{region 'Documentation'}
(*!
<summary>Selects literal stimuli, gates and findings for a named checkpoint.</summary>
*)
{endregion}
METHOD PRIVATE SelectStep : BOOL //! TRUE after selecting a supported script step and its literal expectations; FALSE reports an unknown step.
SelectStep := FALSE;
FIntegerFinding := E_Result.NotEvaluated;
FTextFinding := E_Result.NotEvaluated;
FWideTextFinding := E_Result.NotEvaluated;
FRealFinding := E_Result.NotEvaluated;
FLRealFinding := E_Result.NotEvaluated;
CASE FStep OF
    StepInitialReset:
        FTrace := TraceScalarHistory;
        FResetSubjects := TRUE;
        FSample := 10;
        FTextSample := '10';
        FWideTextSample := "10";
        FRealSample.Value := 10.0;
        FLRealSample.Value := 10.0;
        FIntegerEnable := TRUE;
        FIntegerResult := E_Result.NotEvaluated;
        FIntegerObservation := FALSE;
        FIntegerEvaluation := FALSE;
        FTextEnable := TRUE;
        FTextResult := E_Result.NotEvaluated;
        FTextObservation := FALSE;
        FTextEvaluation := FALSE;
        FWideTextEnable := TRUE;
        FWideTextResult := E_Result.NotEvaluated;
        FWideTextObservation := FALSE;
        FWideTextEvaluation := FALSE;
        FRealEnable := TRUE;
        FRealResult := E_Result.NotEvaluated;
        FRealObservation := FALSE;
        FRealEvaluation := FALSE;
        FLRealEnable := TRUE;
        FLRealResult := E_Result.NotEvaluated;
        FLRealObservation := FALSE;
        FLRealEvaluation := FALSE;
    StepInitialObservation:
        FTrace := TraceScalarHistory;
        FResetSubjects := FALSE;
        FSample := 10;
        FTextSample := '10';
        FWideTextSample := "10";
        FRealSample.Value := 10.0;
        FLRealSample.Value := 10.0;
        FIntegerEnable := TRUE;
        FIntegerResult := E_Result.NotEvaluated;
        FIntegerObservation := TRUE;
        FIntegerEvaluation := FALSE;
        FTextEnable := TRUE;
        FTextResult := E_Result.NotEvaluated;
        FTextObservation := TRUE;
        FTextEvaluation := FALSE;
        FWideTextEnable := TRUE;
        FWideTextResult := E_Result.NotEvaluated;
        FWideTextObservation := TRUE;
        FWideTextEvaluation := FALSE;
        FRealEnable := TRUE;
        FRealResult := E_Result.NotEvaluated;
        FRealObservation := TRUE;
        FRealEvaluation := FALSE;
        FLRealEnable := TRUE;
        FLRealResult := E_Result.NotEvaluated;
        FLRealObservation := TRUE;
        FLRealEvaluation := FALSE;
    StepEqualObservation:
        FTrace := TraceScalarHistory;
        FResetSubjects := FALSE;
        FSample := 10;
        FTextSample := '10';
        FWideTextSample := "10";
        FRealSample.Value := 10.0;
        FLRealSample.Value := 10.0;
        FIntegerEnable := TRUE;
        FIntegerResult := E_Result.Passed;
        FIntegerObservation := TRUE;
        FIntegerEvaluation := TRUE;
        FTextEnable := TRUE;
        FTextResult := E_Result.Passed;
        FTextObservation := TRUE;
        FTextEvaluation := TRUE;
        FWideTextEnable := TRUE;
        FWideTextResult := E_Result.Passed;
        FWideTextObservation := TRUE;
        FWideTextEvaluation := TRUE;
        FRealEnable := TRUE;
        FRealResult := E_Result.Passed;
        FRealObservation := TRUE;
        FRealEvaluation := TRUE;
        FLRealEnable := TRUE;
        FLRealResult := E_Result.Passed;
        FLRealObservation := TRUE;
        FLRealEvaluation := TRUE;
    StepChangedObservation:
        FTrace := TraceScalarHistory;
        FResetSubjects := FALSE;
        FSample := 11;
        FTextSample := '11';
        FWideTextSample := "11";
        FRealSample.Value := 11.0;
        FLRealSample.Value := 11.0;
        FIntegerEnable := TRUE;
        FIntegerResult := E_Result.Failed;
        FIntegerObservation := TRUE;
        FIntegerEvaluation := TRUE;
        FIntegerFinding := E_Result.Failed;
        FTextEnable := TRUE;
        FTextResult := E_Result.Failed;
        FTextObservation := TRUE;
        FTextEvaluation := TRUE;
        FTextFinding := E_Result.Failed;
        FWideTextEnable := TRUE;
        FWideTextResult := E_Result.Failed;
        FWideTextObservation := TRUE;
        FWideTextEvaluation := TRUE;
        FWideTextFinding := E_Result.Failed;
        FRealEnable := TRUE;
        FRealResult := E_Result.Failed;
        FRealObservation := TRUE;
        FRealEvaluation := TRUE;
        FRealFinding := E_Result.Failed;
        FLRealEnable := TRUE;
        FLRealResult := E_Result.Failed;
        FLRealObservation := TRUE;
        FLRealEvaluation := TRUE;
        FLRealFinding := E_Result.Failed;
    StepReturnToInitial:
        FTrace := TraceScalarHistory;
        FResetSubjects := FALSE;
        FSample := 10;
        FTextSample := '10';
        FWideTextSample := "10";
        FRealSample.Value := 10.0;
        FLRealSample.Value := 10.0;
        FIntegerEnable := TRUE;
        FIntegerResult := E_Result.Failed;
        FIntegerObservation := TRUE;
        FIntegerEvaluation := TRUE;
        FTextEnable := TRUE;
        FTextResult := E_Result.Failed;
        FTextObservation := TRUE;
        FTextEvaluation := TRUE;
        FWideTextEnable := TRUE;
        FWideTextResult := E_Result.Failed;
        FWideTextObservation := TRUE;
        FWideTextEvaluation := TRUE;
        FRealEnable := TRUE;
        FRealResult := E_Result.Failed;
        FRealObservation := TRUE;
        FRealEvaluation := TRUE;
        FLRealEnable := TRUE;
        FLRealResult := E_Result.Failed;
        FLRealObservation := TRUE;
        FLRealEvaluation := TRUE;
    StepReenableReset:
        FTrace := TraceReenableBaseline;
        FResetSubjects := TRUE;
        FSample := 10;
        FTextSample := '10';
        FWideTextSample := "10";
        FRealSample.Value := 10.0;
        FLRealSample.Value := 10.0;
        FIntegerEnable := TRUE;
        FIntegerResult := E_Result.NotEvaluated;
        FIntegerObservation := FALSE;
        FIntegerEvaluation := FALSE;
        FTextEnable := TRUE;
        FTextResult := E_Result.NotEvaluated;
        FTextObservation := FALSE;
        FTextEvaluation := FALSE;
        FWideTextEnable := TRUE;
        FWideTextResult := E_Result.NotEvaluated;
        FWideTextObservation := FALSE;
        FWideTextEvaluation := FALSE;
        FRealEnable := TRUE;
        FRealResult := E_Result.NotEvaluated;
        FRealObservation := FALSE;
        FRealEvaluation := FALSE;
        FLRealEnable := TRUE;
        FLRealResult := E_Result.NotEvaluated;
        FLRealObservation := FALSE;
        FLRealEvaluation := FALSE;
    StepReenableBaseline:
        FTrace := TraceReenableBaseline;
        FResetSubjects := FALSE;
        FSample := 10;
        FTextSample := '10';
        FWideTextSample := "10";
        FRealSample.Value := 10.0;
        FLRealSample.Value := 10.0;
        FIntegerEnable := TRUE;
        FIntegerResult := E_Result.NotEvaluated;
        FIntegerObservation := TRUE;
        FIntegerEvaluation := FALSE;
        FTextEnable := TRUE;
        FTextResult := E_Result.NotEvaluated;
        FTextObservation := TRUE;
        FTextEvaluation := FALSE;
        FWideTextEnable := TRUE;
        FWideTextResult := E_Result.NotEvaluated;
        FWideTextObservation := TRUE;
        FWideTextEvaluation := FALSE;
        FRealEnable := TRUE;
        FRealResult := E_Result.NotEvaluated;
        FRealObservation := TRUE;
        FRealEvaluation := FALSE;
        FLRealEnable := TRUE;
        FLRealResult := E_Result.NotEvaluated;
        FLRealObservation := TRUE;
        FLRealEvaluation := FALSE;
    StepBeforeDisable:
        FTrace := TraceReenableBaseline;
        FResetSubjects := FALSE;
        FSample := 10;
        FTextSample := '10';
        FWideTextSample := "10";
        FRealSample.Value := 10.0;
        FLRealSample.Value := 10.0;
        FIntegerEnable := TRUE;
        FIntegerResult := E_Result.Passed;
        FIntegerObservation := TRUE;
        FIntegerEvaluation := TRUE;
        FTextEnable := TRUE;
        FTextResult := E_Result.Passed;
        FTextObservation := TRUE;
        FTextEvaluation := TRUE;
        FWideTextEnable := TRUE;
        FWideTextResult := E_Result.Passed;
        FWideTextObservation := TRUE;
        FWideTextEvaluation := TRUE;
        FRealEnable := TRUE;
        FRealResult := E_Result.Passed;
        FRealObservation := TRUE;
        FRealEvaluation := TRUE;
        FLRealEnable := TRUE;
        FLRealResult := E_Result.Passed;
        FLRealObservation := TRUE;
        FLRealEvaluation := TRUE;
    StepDisabledChange:
        FTrace := TraceReenableBaseline;
        FResetSubjects := FALSE;
        FSample := 20;
        FTextSample := '20';
        FWideTextSample := "20";
        FRealSample.Value := 20.0;
        FLRealSample.Value := 20.0;
        FIntegerEnable := FALSE;
        FIntegerResult := E_Result.Passed;
        FIntegerObservation := FALSE;
        FIntegerEvaluation := FALSE;
        FTextEnable := FALSE;
        FTextResult := E_Result.Passed;
        FTextObservation := FALSE;
        FTextEvaluation := FALSE;
        FWideTextEnable := FALSE;
        FWideTextResult := E_Result.Passed;
        FWideTextObservation := FALSE;
        FWideTextEvaluation := FALSE;
        FRealEnable := FALSE;
        FRealResult := E_Result.Passed;
        FRealObservation := FALSE;
        FRealEvaluation := FALSE;
        FLRealEnable := FALSE;
        FLRealResult := E_Result.Passed;
        FLRealObservation := FALSE;
        FLRealEvaluation := FALSE;
    StepReenabledCapture:
        FTrace := TraceReenableBaseline;
        FResetSubjects := FALSE;
        FSample := 20;
        FTextSample := '20';
        FWideTextSample := "20";
        FRealSample.Value := 20.0;
        FLRealSample.Value := 20.0;
        FIntegerEnable := TRUE;
        FIntegerResult := E_Result.Passed;
        FIntegerObservation := TRUE;
        FIntegerEvaluation := FALSE;
        FTextEnable := TRUE;
        FTextResult := E_Result.Passed;
        FTextObservation := TRUE;
        FTextEvaluation := FALSE;
        FWideTextEnable := TRUE;
        FWideTextResult := E_Result.Passed;
        FWideTextObservation := TRUE;
        FWideTextEvaluation := FALSE;
        FRealEnable := TRUE;
        FRealResult := E_Result.Passed;
        FRealObservation := TRUE;
        FRealEvaluation := FALSE;
        FLRealEnable := TRUE;
        FLRealResult := E_Result.Passed;
        FLRealObservation := TRUE;
        FLRealEvaluation := FALSE;
    StepReenabledComparison:
        FTrace := TraceReenableBaseline;
        FResetSubjects := FALSE;
        FSample := 20;
        FTextSample := '20';
        FWideTextSample := "20";
        FRealSample.Value := 20.0;
        FLRealSample.Value := 20.0;
        FIntegerEnable := TRUE;
        FIntegerResult := E_Result.Passed;
        FIntegerObservation := TRUE;
        FIntegerEvaluation := TRUE;
        FTextEnable := TRUE;
        FTextResult := E_Result.Passed;
        FTextObservation := TRUE;
        FTextEvaluation := TRUE;
        FWideTextEnable := TRUE;
        FWideTextResult := E_Result.Passed;
        FWideTextObservation := TRUE;
        FWideTextEvaluation := TRUE;
        FRealEnable := TRUE;
        FRealResult := E_Result.Passed;
        FRealObservation := TRUE;
        FRealEvaluation := TRUE;
        FLRealEnable := TRUE;
        FLRealResult := E_Result.Passed;
        FLRealObservation := TRUE;
        FLRealEvaluation := TRUE;
    StepResetNewBaseline:
        FTrace := TraceResetBaseline;
        FResetSubjects := TRUE;
        FSample := 30;
        FTextSample := '30';
        FWideTextSample := "30";
        FRealSample.Value := 30.0;
        FLRealSample.Value := 30.0;
        FIntegerEnable := TRUE;
        FIntegerResult := E_Result.NotEvaluated;
        FIntegerObservation := FALSE;
        FIntegerEvaluation := FALSE;
        FTextEnable := TRUE;
        FTextResult := E_Result.NotEvaluated;
        FTextObservation := FALSE;
        FTextEvaluation := FALSE;
        FWideTextEnable := TRUE;
        FWideTextResult := E_Result.NotEvaluated;
        FWideTextObservation := FALSE;
        FWideTextEvaluation := FALSE;
        FRealEnable := TRUE;
        FRealResult := E_Result.NotEvaluated;
        FRealObservation := FALSE;
        FRealEvaluation := FALSE;
        FLRealEnable := TRUE;
        FLRealResult := E_Result.NotEvaluated;
        FLRealObservation := FALSE;
        FLRealEvaluation := FALSE;
    StepNewBaselineCapture:
        FTrace := TraceResetBaseline;
        FResetSubjects := FALSE;
        FSample := 30;
        FTextSample := '30';
        FWideTextSample := "30";
        FRealSample.Value := 30.0;
        FLRealSample.Value := 30.0;
        FIntegerEnable := TRUE;
        FIntegerResult := E_Result.NotEvaluated;
        FIntegerObservation := TRUE;
        FIntegerEvaluation := FALSE;
        FTextEnable := TRUE;
        FTextResult := E_Result.NotEvaluated;
        FTextObservation := TRUE;
        FTextEvaluation := FALSE;
        FWideTextEnable := TRUE;
        FWideTextResult := E_Result.NotEvaluated;
        FWideTextObservation := TRUE;
        FWideTextEvaluation := FALSE;
        FRealEnable := TRUE;
        FRealResult := E_Result.NotEvaluated;
        FRealObservation := TRUE;
        FRealEvaluation := FALSE;
        FLRealEnable := TRUE;
        FLRealResult := E_Result.NotEvaluated;
        FLRealObservation := TRUE;
        FLRealEvaluation := FALSE;
    StepNewBaselineComparison:
        FTrace := TraceResetBaseline;
        FResetSubjects := FALSE;
        FSample := 30;
        FTextSample := '30';
        FWideTextSample := "30";
        FRealSample.Value := 30.0;
        FLRealSample.Value := 30.0;
        FIntegerEnable := TRUE;
        FIntegerResult := E_Result.Passed;
        FIntegerObservation := TRUE;
        FIntegerEvaluation := TRUE;
        FTextEnable := TRUE;
        FTextResult := E_Result.Passed;
        FTextObservation := TRUE;
        FTextEvaluation := TRUE;
        FWideTextEnable := TRUE;
        FWideTextResult := E_Result.Passed;
        FWideTextObservation := TRUE;
        FWideTextEvaluation := TRUE;
        FRealEnable := TRUE;
        FRealResult := E_Result.Passed;
        FRealObservation := TRUE;
        FRealEvaluation := TRUE;
        FLRealEnable := TRUE;
        FLRealResult := E_Result.Passed;
        FLRealObservation := TRUE;
        FLRealEvaluation := TRUE;
    StepNaNReset:
        FTrace := TraceScalarNonFinite;
        FResetSubjects := TRUE;
        FSample := 10;
        FTextSample := '10';
        FWideTextSample := "10";
        FRealSample.Value := 10.0;
        FLRealSample.Value := 10.0;
        FIntegerEnable := FALSE;
        FIntegerResult := E_Result.NotEvaluated;
        FIntegerObservation := FALSE;
        FIntegerEvaluation := FALSE;
        FTextEnable := FALSE;
        FTextResult := E_Result.NotEvaluated;
        FTextObservation := FALSE;
        FTextEvaluation := FALSE;
        FWideTextEnable := FALSE;
        FWideTextResult := E_Result.NotEvaluated;
        FWideTextObservation := FALSE;
        FWideTextEvaluation := FALSE;
        FRealEnable := FALSE;
        FRealResult := E_Result.NotEvaluated;
        FRealObservation := FALSE;
        FRealEvaluation := FALSE;
        FLRealEnable := FALSE;
        FLRealResult := E_Result.NotEvaluated;
        FLRealObservation := FALSE;
        FLRealEvaluation := FALSE;
    StepNaNCapture:
        FTrace := TraceScalarNonFinite;
        FResetSubjects := FALSE;
        FRealSample.Bits := DWORD#16#7FC00000;
        FLRealSample.Bits := LWORD#16#7FF8000000000000;
        FIntegerEnable := FALSE;
        FIntegerResult := E_Result.NotEvaluated;
        FIntegerObservation := FALSE;
        FIntegerEvaluation := FALSE;
        FTextEnable := FALSE;
        FTextResult := E_Result.NotEvaluated;
        FTextObservation := FALSE;
        FTextEvaluation := FALSE;
        FWideTextEnable := FALSE;
        FWideTextResult := E_Result.NotEvaluated;
        FWideTextObservation := FALSE;
        FWideTextEvaluation := FALSE;
        FRealEnable := TRUE;
        FRealResult := E_Result.Error;
        FRealObservation := TRUE;
        FRealEvaluation := FALSE;
        FRealFinding := E_Result.Error;
        FLRealEnable := TRUE;
        FLRealResult := E_Result.Error;
        FLRealObservation := TRUE;
        FLRealEvaluation := FALSE;
        FLRealFinding := E_Result.Error;
    StepNaNRepeated:
        FTrace := TraceScalarNonFinite;
        FResetSubjects := FALSE;
        // The same non-finite input must not produce duplicate findings.
        FIntegerEnable := FALSE;
        FIntegerResult := E_Result.NotEvaluated;
        FIntegerObservation := FALSE;
        FIntegerEvaluation := FALSE;
        FTextEnable := FALSE;
        FTextResult := E_Result.NotEvaluated;
        FTextObservation := FALSE;
        FTextEvaluation := FALSE;
        FWideTextEnable := FALSE;
        FWideTextResult := E_Result.NotEvaluated;
        FWideTextObservation := FALSE;
        FWideTextEvaluation := FALSE;
        FRealEnable := TRUE;
        FRealResult := E_Result.Error;
        FRealObservation := TRUE;
        FRealEvaluation := TRUE;
        FLRealEnable := TRUE;
        FLRealResult := E_Result.Error;
        FLRealObservation := TRUE;
        FLRealEvaluation := TRUE;
    StepPositiveInfinityReset:
        FTrace := TraceScalarNonFinite;
        FResetSubjects := TRUE;
        FSample := 10;
        FTextSample := '10';
        FWideTextSample := "10";
        FRealSample.Value := 10.0;
        FLRealSample.Value := 10.0;
        FIntegerEnable := FALSE;
        FIntegerResult := E_Result.NotEvaluated;
        FIntegerObservation := FALSE;
        FIntegerEvaluation := FALSE;
        FTextEnable := FALSE;
        FTextResult := E_Result.NotEvaluated;
        FTextObservation := FALSE;
        FTextEvaluation := FALSE;
        FWideTextEnable := FALSE;
        FWideTextResult := E_Result.NotEvaluated;
        FWideTextObservation := FALSE;
        FWideTextEvaluation := FALSE;
        FRealEnable := FALSE;
        FRealResult := E_Result.NotEvaluated;
        FRealObservation := FALSE;
        FRealEvaluation := FALSE;
        FLRealEnable := FALSE;
        FLRealResult := E_Result.NotEvaluated;
        FLRealObservation := FALSE;
        FLRealEvaluation := FALSE;
    StepPositiveInfinityCapture:
        FTrace := TraceScalarNonFinite;
        FResetSubjects := FALSE;
        FRealSample.Bits := DWORD#16#7F800000;
        FLRealSample.Bits := LWORD#16#7FF0000000000000;
        FIntegerEnable := FALSE;
        FIntegerResult := E_Result.NotEvaluated;
        FIntegerObservation := FALSE;
        FIntegerEvaluation := FALSE;
        FTextEnable := FALSE;
        FTextResult := E_Result.NotEvaluated;
        FTextObservation := FALSE;
        FTextEvaluation := FALSE;
        FWideTextEnable := FALSE;
        FWideTextResult := E_Result.NotEvaluated;
        FWideTextObservation := FALSE;
        FWideTextEvaluation := FALSE;
        FRealEnable := TRUE;
        FRealResult := E_Result.Error;
        FRealObservation := TRUE;
        FRealEvaluation := FALSE;
        FRealFinding := E_Result.Error;
        FLRealEnable := TRUE;
        FLRealResult := E_Result.Error;
        FLRealObservation := TRUE;
        FLRealEvaluation := FALSE;
        FLRealFinding := E_Result.Error;
    StepPositiveInfinityRepeated:
        FTrace := TraceScalarNonFinite;
        FResetSubjects := FALSE;
        // The same non-finite input must not produce duplicate findings.
        FIntegerEnable := FALSE;
        FIntegerResult := E_Result.NotEvaluated;
        FIntegerObservation := FALSE;
        FIntegerEvaluation := FALSE;
        FTextEnable := FALSE;
        FTextResult := E_Result.NotEvaluated;
        FTextObservation := FALSE;
        FTextEvaluation := FALSE;
        FWideTextEnable := FALSE;
        FWideTextResult := E_Result.NotEvaluated;
        FWideTextObservation := FALSE;
        FWideTextEvaluation := FALSE;
        FRealEnable := TRUE;
        FRealResult := E_Result.Error;
        FRealObservation := TRUE;
        FRealEvaluation := TRUE;
        FLRealEnable := TRUE;
        FLRealResult := E_Result.Error;
        FLRealObservation := TRUE;
        FLRealEvaluation := TRUE;
    StepNegativeInfinityReset:
        FTrace := TraceScalarNonFinite;
        FResetSubjects := TRUE;
        FSample := 10;
        FTextSample := '10';
        FWideTextSample := "10";
        FRealSample.Value := 10.0;
        FLRealSample.Value := 10.0;
        FIntegerEnable := FALSE;
        FIntegerResult := E_Result.NotEvaluated;
        FIntegerObservation := FALSE;
        FIntegerEvaluation := FALSE;
        FTextEnable := FALSE;
        FTextResult := E_Result.NotEvaluated;
        FTextObservation := FALSE;
        FTextEvaluation := FALSE;
        FWideTextEnable := FALSE;
        FWideTextResult := E_Result.NotEvaluated;
        FWideTextObservation := FALSE;
        FWideTextEvaluation := FALSE;
        FRealEnable := FALSE;
        FRealResult := E_Result.NotEvaluated;
        FRealObservation := FALSE;
        FRealEvaluation := FALSE;
        FLRealEnable := FALSE;
        FLRealResult := E_Result.NotEvaluated;
        FLRealObservation := FALSE;
        FLRealEvaluation := FALSE;
    StepNegativeInfinityCapture:
        FTrace := TraceScalarNonFinite;
        FResetSubjects := FALSE;
        FRealSample.Bits := DWORD#16#FF800000;
        FLRealSample.Bits := LWORD#16#FFF0000000000000;
        FIntegerEnable := FALSE;
        FIntegerResult := E_Result.NotEvaluated;
        FIntegerObservation := FALSE;
        FIntegerEvaluation := FALSE;
        FTextEnable := FALSE;
        FTextResult := E_Result.NotEvaluated;
        FTextObservation := FALSE;
        FTextEvaluation := FALSE;
        FWideTextEnable := FALSE;
        FWideTextResult := E_Result.NotEvaluated;
        FWideTextObservation := FALSE;
        FWideTextEvaluation := FALSE;
        FRealEnable := TRUE;
        FRealResult := E_Result.Error;
        FRealObservation := TRUE;
        FRealEvaluation := FALSE;
        FRealFinding := E_Result.Error;
        FLRealEnable := TRUE;
        FLRealResult := E_Result.Error;
        FLRealObservation := TRUE;
        FLRealEvaluation := FALSE;
        FLRealFinding := E_Result.Error;
    StepNegativeInfinityRepeated:
        FTrace := TraceScalarNonFinite;
        FResetSubjects := FALSE;
        // The same non-finite input must not produce duplicate findings.
        FIntegerEnable := FALSE;
        FIntegerResult := E_Result.NotEvaluated;
        FIntegerObservation := FALSE;
        FIntegerEvaluation := FALSE;
        FTextEnable := FALSE;
        FTextResult := E_Result.NotEvaluated;
        FTextObservation := FALSE;
        FTextEvaluation := FALSE;
        FWideTextEnable := FALSE;
        FWideTextResult := E_Result.NotEvaluated;
        FWideTextObservation := FALSE;
        FWideTextEvaluation := FALSE;
        FRealEnable := TRUE;
        FRealResult := E_Result.Error;
        FRealObservation := TRUE;
        FRealEvaluation := TRUE;
        FLRealEnable := TRUE;
        FLRealResult := E_Result.Error;
        FLRealObservation := TRUE;
        FLRealEvaluation := TRUE;
ELSE
    Error(Message := 'Unknown observation checkpoint.');
    RETURN;
END_CASE;
SelectStep := TRUE;
END_METHOD

END_FUNCTION_BLOCK

// ---- Framework/Assertions/POU/BasicTypes/DInt/AssertNoValueChange_DInt.TcPOU
{region 'Documentation'}
(*!
<summary>Check equality between consecutive active observations.</summary>
<description>

The first active observation establishes a baseline without deciding a result. Disabling
observation invalidates that baseline, not the held Result. Re-enabling first establishes a new
baseline; Reset clears history.

ObserveFirstCycle FALSE delays the first observation by one enabled call.

</description>
*)
{endregion}
FUNCTION_BLOCK AssertNoValueChange_DInt EXTENDS AssertionBase
VAR_INPUT
    IN : DINT; //! Actual value to observe.
END_VAR
VAR
    FINPrevious : DINT;
    FObservationPrevious : BOOL;
    FEvaluationActive : BOOL;
END_VAR

SUPER^();

{region 'Documentation'}
(*!
<summary>Observe the current value before evaluating a change against the previous observation.</summary>
*)
{endregion}
METHOD PROTECTED Assert
VAR
    PreviousValue : DINT;
    Message : STRING(GVL_Constants.MessageLength);
    PreviousText : STRING(GVL_Constants.AssertionValueLength);
    ActualText : STRING(GVL_Constants.AssertionValueLength);
END_VAR
FEvaluationActive := ObservationActive AND FObservationPrevious;
FObservationPrevious := ObservationActive;

IF NOT ObservationActive THEN
    RETURN;
END_IF;

PreviousValue := FINPrevious;
FINPrevious := IN;

IF NOT EvaluationActive THEN
    RETURN;
END_IF;

IF Result = E_Result.Error THEN
    RETURN;
END_IF;

IF Result = E_Result.Failed THEN
    RETURN;
END_IF;

IF IN <> PreviousValue THEN
    PreviousText := DINT_TO_STRING(PreviousValue);
    ActualText := DINT_TO_STRING(IN);
    Message := CONCAT('Assertion failed: value changed unexpectedly. Previous = ',
        PreviousText);
    Message := CONCAT(Message, ', Actual = ');
    Message := CONCAT(Message, ActualText);
    Message := CONCAT(Message, '.');
    Fail(Message := Message);
    RETURN;
END_IF;

Pass();
END_METHOD

{region 'Documentation'}
(*!
<summary>Current/last call has an active observation and a preceding observation
baseline.</summary>
*)
{endregion}
{attribute 'monitoring' := 'call'}
PROPERTY PUBLIC EvaluationActive : BOOL //! Current/last call has an active observation and a preceding observation baseline.
GET // PUBLIC
EvaluationActive := FEvaluationActive;
END_GET
END_PROPERTY

{region 'Documentation'}
(*!
<summary>Clear observation history and the current evaluation gate.</summary>
*)
{endregion}
METHOD PROTECTED ResetAssertion
FINPrevious := 0;
FObservationPrevious := FALSE;
FEvaluationActive := FALSE;
END_METHOD

END_FUNCTION_BLOCK

// ---- Framework/Assertions/POU/BasicTypes/LReal/AssertNoValueChange_LReal.TcPOU
{region 'Documentation'}
(*!
<summary>Check equality between consecutive active observations.</summary>
<description>

The first active observation establishes a baseline without deciding a result. Disabling
observation invalidates that baseline, not the held Result. Re-enabling first establishes a new
baseline; Reset clears history.

ObserveFirstCycle FALSE delays the first observation by one enabled call.

NaN or either infinity reports Error on an active observation, including baseline
capture; finite values compare exactly.

Numeric diagnostics use the formatter's default six significant digits; rounding affects
the message only, not the comparison.

</description>
*)
{endregion}
FUNCTION_BLOCK AssertNoValueChange_LReal EXTENDS AssertionBase
VAR_INPUT
    IN : LREAL; //! Actual value to observe.
END_VAR
VAR
    FINPrevious : LREAL;
    FObservationPrevious : BOOL;
    FEvaluationActive : BOOL;
END_VAR

SUPER^();

{region 'Documentation'}
(*!
<summary>Observe the current value before evaluating a change against the previous observation.</summary>
*)
{endregion}
METHOD PROTECTED Assert
VAR
    PreviousValue : LREAL;
    Message : STRING(GVL_Constants.MessageLength);
    PreviousText : STRING(GVL_Constants.AssertionValueLength);
    ActualText : STRING(GVL_Constants.AssertionValueLength);
END_VAR
FEvaluationActive := ObservationActive AND FObservationPrevious;
FObservationPrevious := ObservationActive;

IF NOT ObservationActive THEN
    RETURN;
END_IF;

PreviousValue := FINPrevious;
FINPrevious := IN;

IF Result = E_Result.Error THEN
    RETURN;
END_IF;

IF NOT Tc2_Utilities.LrealIsFinite(x := IN) THEN
    Error(Message := 'Assertion error: IN must be finite.');
    RETURN;
END_IF;

IF NOT EvaluationActive THEN
    RETURN;
END_IF;

IF Result = E_Result.Failed THEN
    RETURN;
END_IF;

IF IN <> PreviousValue THEN
    PreviousText := CreateAssertionTextValue_LReal(Value := PreviousValue);
    ActualText := CreateAssertionTextValue_LReal(Value := IN);
    Message := CONCAT('Assertion failed: value changed unexpectedly. Previous = ',
        PreviousText);
    Message := CONCAT(Message, ', Actual = ');
    Message := CONCAT(Message, ActualText);
    Message := CONCAT(Message, '.');
    Fail(Message := Message);
    RETURN;
END_IF;

Pass();
END_METHOD

{region 'Documentation'}
(*!
<summary>Current/last call has an active observation and a preceding observation
baseline.</summary>
*)
{endregion}
{attribute 'monitoring' := 'call'}
PROPERTY PUBLIC EvaluationActive : BOOL //! Current/last call has an active observation and a preceding observation baseline.
GET // PUBLIC
EvaluationActive := FEvaluationActive;
END_GET
END_PROPERTY

{region 'Documentation'}
(*!
<summary>Clear observation history and the current evaluation gate.</summary>
*)
{endregion}
METHOD PROTECTED ResetAssertion
FINPrevious := 0.0;
FObservationPrevious := FALSE;
FEvaluationActive := FALSE;
END_METHOD

END_FUNCTION_BLOCK

// ---- SelfTests/TestCases/TestSuite_AssertionObservation/Test_AssertionArraySnapshot.TcPOU
{region 'Documentation'}
(*!
<summary>Checks retained DINT array snapshots, independent bounds and delayed observation.</summary>
<description>
IN[-2..1] selects [-1..0], while Memory[5..7] stores two values and an untouched
tail sentinel. Disable never replaces the snapshot. Reset invalidates it without
clearing Memory; ObserveFirstCycle=FALSE delays capture until the second enabled
call. Literal memory checks distinguish fixed snapshots from rolling history.
Each named step calls each subject once and checks public gates, result and local
findings before advancing in the next cycle. Outer Assertions collect checkpoints
per trace; subjects never contribute their intentional failures to the test result.
FirstFailedStep retains the first mismatch. No timed stimulus or expected-result
algorithm is used.
</description>
*)
{endregion}
FUNCTION_BLOCK Test_AssertionArraySnapshot EXTENDS TestCaseBase
VAR
    FImmediate : AssertArrayNoValueChange_DInt;
    FDelayed : AssertArrayNoValueChange_DInt;
    FInput : ARRAY[-2..1] OF DINT;
    FImmediateMemory : ARRAY[5..7] OF DINT;
    FDelayedMemory : ARRAY[5..7] OF DINT;
    FExpectedImmediateFirst : DINT;
    FExpectedImmediateSecond : DINT;
    FExpectedDelayedFirst : DINT;
    FExpectedDelayedSecond : DINT;
    FCapture : EventBuffer;
    FEvents : ARRAY[1..CaptureLength] OF ST_Event;
    FCaptureFifo : ST_FifoStatus;
    FCaptureStatus : ST_EventBufferStatus;
    FSetupValid : BOOL;
    FStep : UINT;
    FTrace : UINT;
    FFirstFailedStep : UINT;
    FChecked : BOOL;
    FObservationReady : BOOL;
    FStepMatches : BOOL;
    FResultsMatch : BOOL;
    FActivityMatches : BOOL;
    FFindingsMatch : BOOL;
    FMemoryMatches : BOOL;
    FResetSubjects : BOOL;
    FImmediateEnable : BOOL;
    FImmediateResult : E_Result;
    FImmediateObservation : BOOL;
    FImmediateEvaluation : BOOL;
    FImmediateFinding : E_Result;
    FDelayedEnable : BOOL;
    FDelayedResult : E_Result;
    FDelayedObservation : BOOL;
    FDelayedEvaluation : BOOL;
    FDelayedFinding : E_Result;
    FFixedSnapshot : AssertTrue;
    FRetainedOnReenable : AssertTrue;
    FRecaptureAfterReset : AssertTrue;
END_VAR
VAR CONSTANT
    CaptureLength : UINT := 8;
    StepResetSnapshot : UINT := 1;
    StepFirstObservation : UINT := 2;
    StepDelayedCapture : UINT := 3;
    StepEqualSnapshot : UINT := 4;
    StepDivergence : UINT := 5;
    StepReturnToSnapshot : UINT := 6;
    StepResetForReenable : UINT := 7;
    StepReenableTraceCapture : UINT := 8;
    StepReenableTraceDelayedCapture : UINT := 9;
    StepReenableTracePassed : UINT := 10;
    StepDisabledChange : UINT := 11;
    StepReenableHistory : UINT := 12;
    StepReenableComparison : UINT := 13;
    StepReenableDelayedComparison : UINT := 14;
    StepResetKeepsMemory : UINT := 15;
    StepNewSnapshot : UINT := 16;
    StepNewDelayedSnapshot : UINT := 17;
    StepNewSnapshotMatches : UINT := 18;
    LastStep : UINT := StepNewSnapshotMatches;
    TraceFixedSnapshot : UINT := 1;
    TraceRetainedOnReenable : UINT := 2;
    TraceRecaptureAfterReset : UINT := 3;
END_VAR

SUPER^();

{region 'Documentation'}
(*!
<summary>Aggregates only the outer checks, not the intentionally failing subjects.</summary>
*)
{endregion}
METHOD PROTECTED AggregateResults
VAR_INPUT
    Aggregator : I_ResultAggregator; //! Borrowed result sink owned by the outer Test Case; add this test's checking Assertions without resetting or retaining the sink.
END_VAR
Aggregator.AddProvider(Provider := FFixedSnapshot);
Aggregator.AddProvider(Provider := FRetainedOnReenable);
Aggregator.AddProvider(Provider := FRecaptureAfterReset);
END_METHOD

{region 'Documentation'}
(*!
<summary>Calls each production subject with stable bindings and the selected stimulus.</summary>
*)
{endregion}
METHOD PRIVATE CallSubjects
FImmediate(Enable := FImmediateEnable,
    State := E_State.Running,
    StartIndex := -1,
    Length := 2,
    IN := FInput,
    Memory := FImmediateMemory);
FDelayed(Enable := FDelayedEnable,
    State := E_State.Running,
    StartIndex := -1,
    Length := 2,
    IN := FInput,
    Memory := FDelayedMemory);
END_METHOD

{region 'Documentation'}
(*!
<summary>Checks finding order, identities and exact count without retaining prior events.</summary>
*)
{endregion}
METHOD PRIVATE CheckFindings
VAR
    Index : UINT;
    FindingMatches : BOOL;
END_VAR
Index := 1;
FFindingsMatch := TRUE;
IF FImmediateFinding <> E_Result.NotEvaluated THEN
    FindingMatches := IsFindingValid(Index := Index,
        ExpectedName := FImmediate.Name,
        ExpectedResult := FImmediateFinding);
    FFindingsMatch := FFindingsMatch AND FindingMatches;
    Index := Index + 1;
END_IF;
IF FDelayedFinding <> E_Result.NotEvaluated THEN
    FindingMatches := IsFindingValid(Index := Index,
        ExpectedName := FDelayed.Name,
        ExpectedResult := FDelayedFinding);
    FFindingsMatch := FFindingsMatch AND FindingMatches;
    Index := Index + 1;
END_IF;
FFindingsMatch := FFindingsMatch
    AND (FCaptureStatus.SequenceId = UINT_TO_UDINT(Index - 1))
    AND (FCaptureStatus.LostEventCount = 0);
END_METHOD

{region 'Documentation'}
(*!
<summary>Rejects an incomplete capture or subject setup.</summary>
*)
{endregion}
METHOD PROTECTED CheckInitialization : BOOL //! TRUE when the inherited initialization check and this concrete fixture check both accept the setup.
CheckInitialization := SUPER^.CheckInitialization();
IF NOT CheckInitialization THEN
    RETURN;
END_IF;

CheckInitialization := FSetupValid
    AND FFixedSnapshot.IsInitialized
    AND FRetainedOnReenable.IsInitialized
    AND FRecaptureAfterReset.IsInitialized;
IF NOT CheckInitialization THEN
    EventPublisher.PublishEvent(Event := CreateFrameworkEvent(Name := Name,
        ResourceName := '',
        State := State,
        Severity := E_EventSeverity.Error,
        Message := 'Observation selftest setup failed.'));
END_IF;
END_METHOD

{region 'Documentation'}
(*!
<summary>Checks the selected snapshot and untouched sentinels.</summary>
*)
{endregion}
METHOD PRIVATE CheckMemory
FMemoryMatches := (FImmediateMemory[5] = FExpectedImmediateFirst)
    AND (FImmediateMemory[6] = FExpectedImmediateSecond)
    AND (FDelayedMemory[5] = FExpectedDelayedFirst)
    AND (FDelayedMemory[6] = FExpectedDelayedSecond)
    AND (FImmediateMemory[7] = -999)
    AND (FDelayedMemory[7] = -999)
    AND (FInput[-2] = -100)
    AND (FInput[1] = 100);
END_METHOD

{region 'Documentation'}
(*!
<summary>Checks literal result and observation/evaluation expectations.</summary>
*)
{endregion}
METHOD PRIVATE CheckResults
FResultsMatch := (FImmediate.Result = FImmediateResult)
    AND (FDelayed.Result = FDelayedResult);
FActivityMatches := (FImmediate.Enabled = FImmediateEnable)
    AND (FImmediate.ObservationActive = FImmediateObservation)
    AND (FImmediate.EvaluationActive = FImmediateEvaluation)
    AND (FDelayed.Enabled = FDelayedEnable)
    AND (FDelayed.ObservationActive = FDelayedObservation)
    AND (FDelayed.EvaluationActive = FDelayedEvaluation);
END_METHOD

{region 'Documentation'}
(*!
<summary>Initializes outer checks and isolates intentional subject findings.</summary>
*)
{endregion}
METHOD PROTECTED Configure
VAR
    Initialized : BOOL;
END_VAR
FPreparationStateCount := 0;
FTestStateCount := 1;
FFixedSnapshot.Initialize(Parent := THIS^,
    AssertionName := 'FixedSnapshot');
FRetainedOnReenable.Initialize(Parent := THIS^,
    AssertionName := 'RetainedOnReenable');
FRecaptureAfterReset.Initialize(Parent := THIS^,
    AssertionName := 'RecaptureAfterReset');
FSetupValid := FCapture.Initialize(Buffer := FEvents,
    FifoControl := FCaptureFifo,
    Status := FCaptureStatus);
FImmediate.BindPublisher(Publisher := FCapture);
Initialized := FImmediate.Initialize(Parent := THIS^,
    AssertionName := 'Immediate',
    ObserveFirstCycle := TRUE);
FSetupValid := FSetupValid AND Initialized;
FDelayed.BindPublisher(Publisher := FCapture);
Initialized := FDelayed.Initialize(Parent := THIS^,
    AssertionName := 'Delayed',
    ObserveFirstCycle := FALSE);
FSetupValid := FSetupValid AND Initialized;
END_METHOD

{region 'Documentation'}
(*!
<summary>Checks one expected Failed or Error finding from the bounded local capture.</summary>
*)
{endregion}
METHOD PRIVATE IsFindingValid : BOOL //! TRUE when the selected captured finding satisfies the scenario metadata and diagnostic checks.
VAR_INPUT
    Index : UINT; //! One-based index in the retained isolated event capture.
    ExpectedName : STRING(GVL_Constants.NameLength); //! Independently authored Assertion name expected in the selected finding.
    ExpectedResult : E_Result; //! Independently authored finding result.
END_VAR
IsFindingValid := (FEvents[Index].SequenceId = UINT_TO_UDINT(Index))
    AND (FEvents[Index].Name = ExpectedName)
    AND (FEvents[Index].OwnerScope = E_OwnerScope.Assertion)
    AND (FEvents[Index].EventType = E_EventType.Result)
    AND (FEvents[Index].State = E_State.Running)
    AND (FEvents[Index].Result = ExpectedResult)
    AND (FEvents[Index].Message <> '');
END_METHOD

{region 'Documentation'}
(*!
<summary>Completes abort without asynchronous resources.</summary>
*)
{endregion}
METHOD PROTECTED ProcessAbort
VAR_INPUT
    Enable : BOOL; //! Phase permission supplied by the owning Test Case; FALSE does not authorize progression, while observation may continue.
END_VAR
IF Enable THEN
    CompleteAbort();
END_IF;
END_METHOD

{region 'Documentation'}
(*!
<summary>Checks this checkpoint before the next cycle advances the trace.</summary>
*)
{endregion}
METHOD PROTECTED ProcessAssertions
VAR_INPUT
    Enable : BOOL; //! Phase permission supplied by the owning Test Case; FALSE does not authorize progression, while observation may continue.
END_VAR
VAR
    Check : BOOL;
END_VAR
Check := Enable AND FObservationReady;
FFixedSnapshot(Enable := Check AND (FTrace = TraceFixedSnapshot),
    State := State,
    IN := FStepMatches);
FRetainedOnReenable(Enable := Check AND (FTrace = TraceRetainedOnReenable),
    State := State,
    IN := FStepMatches);
FRecaptureAfterReset(Enable := Check AND (FTrace = TraceRecaptureAfterReset),
    State := State,
    IN := FStepMatches);
IF Check THEN
    FChecked := TRUE;
END_IF;
END_METHOD

{region 'Documentation'}
(*!
<summary>No Preparation phase is required.</summary>
*)
{endregion}
METHOD PROTECTED ProcessPreparations
VAR_INPUT
    // SA0033: Required hook; this test has no Preparation phase.
    {attribute 'analysis' := '-33'}
    Enable : BOOL; //! Phase permission supplied by the owning Test Case; FALSE does not authorize progression, while observation may continue.
END_VAR
END_METHOD

{region 'Documentation'}
(*!
<summary>Resets checkpoint bookkeeping and queues each subject reset.</summary>
*)
{endregion}
METHOD PROTECTED ProcessReset
FStep := StepResetSnapshot;
FTrace := 0;
FFirstFailedStep := 0;
FChecked := FALSE;
FObservationReady := FALSE;
FCapture.Reset();
ResetSubjects();
FFixedSnapshot.Reset();
FRetainedOnReenable.Reset();
FRecaptureAfterReset.Reset();
CompleteReset();
END_METHOD

{region 'Documentation'}
(*!
<summary>Executes exactly one named checkpoint per active PLC cycle.</summary>
*)
{endregion}
METHOD PROTECTED ProcessTests
VAR_INPUT
    Enable : BOOL; //! Phase permission supplied by the owning Test Case; FALSE does not authorize progression, while observation may continue.
END_VAR
IF NOT Enable THEN
    RETURN;
END_IF;

IF FChecked THEN
    FChecked := FALSE;
    FObservationReady := FALSE;
    IF FStep = LastStep THEN
        CompleteTests();
        RETURN;
    END_IF;
    FStep := FStep + 1;
END_IF;

IF NOT SelectStep() THEN
    RETURN;
END_IF;
FCapture.Reset();
IF FResetSubjects THEN
    ResetSubjects();
END_IF;
CallSubjects();
CheckResults();
CheckMemory();
CheckFindings();
FStepMatches := FResultsMatch AND FActivityMatches AND FMemoryMatches AND FFindingsMatch;
IF NOT FStepMatches AND (FFirstFailedStep = 0) THEN
    FFirstFailedStep := FStep;
END_IF;
FObservationReady := TRUE;
END_METHOD

{region 'Documentation'}
(*!
<summary>Queues subject reset; the next bound call consumes it.</summary>
*)
{endregion}
METHOD PRIVATE ResetSubjects
FImmediate.Reset();
FDelayed.Reset();
END_METHOD

{region 'Documentation'}
(*!
<summary>Selects literal stimuli, gates and findings for a named checkpoint.</summary>
*)
{endregion}
METHOD PRIVATE SelectStep : BOOL //! TRUE after selecting a supported script step and its literal expectations; FALSE reports an unknown step.
SelectStep := FALSE;
FImmediateFinding := E_Result.NotEvaluated;
FDelayedFinding := E_Result.NotEvaluated;
CASE FStep OF
    StepResetSnapshot:
        FTrace := TraceFixedSnapshot;
        FResetSubjects := TRUE;
        FInput[-2] := -100;
        FInput[-1] := 10;
        FInput[0] := 20;
        FInput[1] := 100;
        FExpectedImmediateFirst := -777;
        FExpectedImmediateSecond := -888;
        FExpectedDelayedFirst := -777;
        FExpectedDelayedSecond := -888;
        FImmediateMemory[5] := -777;
        FImmediateMemory[6] := -888;
        FImmediateMemory[7] := -999;
        FDelayedMemory[5] := -777;
        FDelayedMemory[6] := -888;
        FDelayedMemory[7] := -999;
        FImmediateEnable := TRUE;
        FImmediateResult := E_Result.NotEvaluated;
        FImmediateObservation := FALSE;
        FImmediateEvaluation := FALSE;
        FDelayedEnable := TRUE;
        FDelayedResult := E_Result.NotEvaluated;
        FDelayedObservation := FALSE;
        FDelayedEvaluation := FALSE;
    StepFirstObservation:
        FTrace := TraceFixedSnapshot;
        FResetSubjects := FALSE;
        FInput[-2] := -100;
        FInput[-1] := 10;
        FInput[0] := 20;
        FInput[1] := 100;
        FExpectedImmediateFirst := 10;
        FExpectedImmediateSecond := 20;
        FExpectedDelayedFirst := -777;
        FExpectedDelayedSecond := -888;
        FImmediateEnable := TRUE;
        FImmediateResult := E_Result.NotEvaluated;
        FImmediateObservation := TRUE;
        FImmediateEvaluation := FALSE;
        FDelayedEnable := TRUE;
        FDelayedResult := E_Result.NotEvaluated;
        FDelayedObservation := FALSE;
        FDelayedEvaluation := FALSE;
    StepDelayedCapture:
        FTrace := TraceFixedSnapshot;
        FResetSubjects := FALSE;
        FInput[-2] := -100;
        FInput[-1] := 10;
        FInput[0] := 20;
        FInput[1] := 100;
        FExpectedImmediateFirst := 10;
        FExpectedImmediateSecond := 20;
        FExpectedDelayedFirst := 10;
        FExpectedDelayedSecond := 20;
        FImmediateEnable := TRUE;
        FImmediateResult := E_Result.Passed;
        FImmediateObservation := TRUE;
        FImmediateEvaluation := TRUE;
        FDelayedEnable := TRUE;
        FDelayedResult := E_Result.NotEvaluated;
        FDelayedObservation := TRUE;
        FDelayedEvaluation := FALSE;
    StepEqualSnapshot:
        FTrace := TraceFixedSnapshot;
        FResetSubjects := FALSE;
        FInput[-2] := -100;
        FInput[-1] := 10;
        FInput[0] := 20;
        FInput[1] := 100;
        FExpectedImmediateFirst := 10;
        FExpectedImmediateSecond := 20;
        FExpectedDelayedFirst := 10;
        FExpectedDelayedSecond := 20;
        FImmediateEnable := TRUE;
        FImmediateResult := E_Result.Passed;
        FImmediateObservation := TRUE;
        FImmediateEvaluation := TRUE;
        FDelayedEnable := TRUE;
        FDelayedResult := E_Result.Passed;
        FDelayedObservation := TRUE;
        FDelayedEvaluation := TRUE;
    StepDivergence:
        FTrace := TraceFixedSnapshot;
        FResetSubjects := FALSE;
        FInput[-2] := -100;
        FInput[-1] := 11;
        FInput[0] := 20;
        FInput[1] := 100;
        FExpectedImmediateFirst := 10;
        FExpectedImmediateSecond := 20;
        FExpectedDelayedFirst := 10;
        FExpectedDelayedSecond := 20;
        FImmediateEnable := TRUE;
        FImmediateResult := E_Result.Failed;
        FImmediateObservation := TRUE;
        FImmediateEvaluation := TRUE;
        FImmediateFinding := E_Result.Failed;
        FDelayedEnable := TRUE;
        FDelayedResult := E_Result.Failed;
        FDelayedObservation := TRUE;
        FDelayedEvaluation := TRUE;
        FDelayedFinding := E_Result.Failed;
    StepReturnToSnapshot:
        FTrace := TraceFixedSnapshot;
        FResetSubjects := FALSE;
        FInput[-2] := -100;
        FInput[-1] := 10;
        FInput[0] := 20;
        FInput[1] := 100;
        FExpectedImmediateFirst := 10;
        FExpectedImmediateSecond := 20;
        FExpectedDelayedFirst := 10;
        FExpectedDelayedSecond := 20;
        FImmediateEnable := TRUE;
        FImmediateResult := E_Result.Failed;
        FImmediateObservation := TRUE;
        FImmediateEvaluation := TRUE;
        FDelayedEnable := TRUE;
        FDelayedResult := E_Result.Failed;
        FDelayedObservation := TRUE;
        FDelayedEvaluation := TRUE;
    StepResetForReenable:
        FTrace := TraceRetainedOnReenable;
        FResetSubjects := TRUE;
        FInput[-2] := -100;
        FInput[-1] := 10;
        FInput[0] := 20;
        FInput[1] := 100;
        FExpectedImmediateFirst := 10;
        FExpectedImmediateSecond := 20;
        FExpectedDelayedFirst := 10;
        FExpectedDelayedSecond := 20;
        FImmediateEnable := TRUE;
        FImmediateResult := E_Result.NotEvaluated;
        FImmediateObservation := FALSE;
        FImmediateEvaluation := FALSE;
        FDelayedEnable := TRUE;
        FDelayedResult := E_Result.NotEvaluated;
        FDelayedObservation := FALSE;
        FDelayedEvaluation := FALSE;
    StepReenableTraceCapture:
        FTrace := TraceRetainedOnReenable;
        FResetSubjects := FALSE;
        FInput[-2] := -100;
        FInput[-1] := 10;
        FInput[0] := 20;
        FInput[1] := 100;
        FExpectedImmediateFirst := 10;
        FExpectedImmediateSecond := 20;
        FExpectedDelayedFirst := 10;
        FExpectedDelayedSecond := 20;
        FImmediateEnable := TRUE;
        FImmediateResult := E_Result.NotEvaluated;
        FImmediateObservation := TRUE;
        FImmediateEvaluation := FALSE;
        FDelayedEnable := TRUE;
        FDelayedResult := E_Result.NotEvaluated;
        FDelayedObservation := FALSE;
        FDelayedEvaluation := FALSE;
    StepReenableTraceDelayedCapture:
        FTrace := TraceRetainedOnReenable;
        FResetSubjects := FALSE;
        FInput[-2] := -100;
        FInput[-1] := 10;
        FInput[0] := 20;
        FInput[1] := 100;
        FExpectedImmediateFirst := 10;
        FExpectedImmediateSecond := 20;
        FExpectedDelayedFirst := 10;
        FExpectedDelayedSecond := 20;
        FImmediateEnable := TRUE;
        FImmediateResult := E_Result.Passed;
        FImmediateObservation := TRUE;
        FImmediateEvaluation := TRUE;
        FDelayedEnable := TRUE;
        FDelayedResult := E_Result.NotEvaluated;
        FDelayedObservation := TRUE;
        FDelayedEvaluation := FALSE;
    StepReenableTracePassed:
        FTrace := TraceRetainedOnReenable;
        FResetSubjects := FALSE;
        FInput[-2] := -100;
        FInput[-1] := 10;
        FInput[0] := 20;
        FInput[1] := 100;
        FExpectedImmediateFirst := 10;
        FExpectedImmediateSecond := 20;
        FExpectedDelayedFirst := 10;
        FExpectedDelayedSecond := 20;
        FImmediateEnable := TRUE;
        FImmediateResult := E_Result.Passed;
        FImmediateObservation := TRUE;
        FImmediateEvaluation := TRUE;
        FDelayedEnable := TRUE;
        FDelayedResult := E_Result.Passed;
        FDelayedObservation := TRUE;
        FDelayedEvaluation := TRUE;
    StepDisabledChange:
        FTrace := TraceRetainedOnReenable;
        FResetSubjects := FALSE;
        FInput[-2] := -100;
        FInput[-1] := 30;
        FInput[0] := 20;
        FInput[1] := 100;
        FExpectedImmediateFirst := 10;
        FExpectedImmediateSecond := 20;
        FExpectedDelayedFirst := 10;
        FExpectedDelayedSecond := 20;
        FImmediateEnable := FALSE;
        FImmediateResult := E_Result.Passed;
        FImmediateObservation := FALSE;
        FImmediateEvaluation := FALSE;
        FDelayedEnable := FALSE;
        FDelayedResult := E_Result.Passed;
        FDelayedObservation := FALSE;
        FDelayedEvaluation := FALSE;
    StepReenableHistory:
        FTrace := TraceRetainedOnReenable;
        FResetSubjects := FALSE;
        FInput[-2] := -100;
        FInput[-1] := 30;
        FInput[0] := 20;
        FInput[1] := 100;
        FExpectedImmediateFirst := 10;
        FExpectedImmediateSecond := 20;
        FExpectedDelayedFirst := 10;
        FExpectedDelayedSecond := 20;
        FImmediateEnable := TRUE;
        FImmediateResult := E_Result.Passed;
        FImmediateObservation := TRUE;
        FImmediateEvaluation := FALSE;
        FDelayedEnable := TRUE;
        FDelayedResult := E_Result.Passed;
        FDelayedObservation := FALSE;
        FDelayedEvaluation := FALSE;
    StepReenableComparison:
        FTrace := TraceRetainedOnReenable;
        FResetSubjects := FALSE;
        FInput[-2] := -100;
        FInput[-1] := 30;
        FInput[0] := 20;
        FInput[1] := 100;
        FExpectedImmediateFirst := 10;
        FExpectedImmediateSecond := 20;
        FExpectedDelayedFirst := 10;
        FExpectedDelayedSecond := 20;
        FImmediateEnable := TRUE;
        FImmediateResult := E_Result.Failed;
        FImmediateObservation := TRUE;
        FImmediateEvaluation := TRUE;
        FImmediateFinding := E_Result.Failed;
        FDelayedEnable := TRUE;
        FDelayedResult := E_Result.Passed;
        FDelayedObservation := TRUE;
        FDelayedEvaluation := FALSE;
    StepReenableDelayedComparison:
        FTrace := TraceRetainedOnReenable;
        FResetSubjects := FALSE;
        FInput[-2] := -100;
        FInput[-1] := 30;
        FInput[0] := 20;
        FInput[1] := 100;
        FExpectedImmediateFirst := 10;
        FExpectedImmediateSecond := 20;
        FExpectedDelayedFirst := 10;
        FExpectedDelayedSecond := 20;
        FImmediateEnable := TRUE;
        FImmediateResult := E_Result.Failed;
        FImmediateObservation := TRUE;
        FImmediateEvaluation := TRUE;
        FDelayedEnable := TRUE;
        FDelayedResult := E_Result.Failed;
        FDelayedObservation := TRUE;
        FDelayedEvaluation := TRUE;
        FDelayedFinding := E_Result.Failed;
    StepResetKeepsMemory:
        FTrace := TraceRecaptureAfterReset;
        FResetSubjects := TRUE;
        FInput[-2] := -100;
        FInput[-1] := 40;
        FInput[0] := 20;
        FInput[1] := 100;
        FExpectedImmediateFirst := 10;
        FExpectedImmediateSecond := 20;
        FExpectedDelayedFirst := 10;
        FExpectedDelayedSecond := 20;
        FImmediateEnable := TRUE;
        FImmediateResult := E_Result.NotEvaluated;
        FImmediateObservation := FALSE;
        FImmediateEvaluation := FALSE;
        FDelayedEnable := TRUE;
        FDelayedResult := E_Result.NotEvaluated;
        FDelayedObservation := FALSE;
        FDelayedEvaluation := FALSE;
    StepNewSnapshot:
        FTrace := TraceRecaptureAfterReset;
        FResetSubjects := FALSE;
        FInput[-2] := -100;
        FInput[-1] := 40;
        FInput[0] := 20;
        FInput[1] := 100;
        FExpectedImmediateFirst := 40;
        FExpectedImmediateSecond := 20;
        FExpectedDelayedFirst := 10;
        FExpectedDelayedSecond := 20;
        FImmediateEnable := TRUE;
        FImmediateResult := E_Result.NotEvaluated;
        FImmediateObservation := TRUE;
        FImmediateEvaluation := FALSE;
        FDelayedEnable := TRUE;
        FDelayedResult := E_Result.NotEvaluated;
        FDelayedObservation := FALSE;
        FDelayedEvaluation := FALSE;
    StepNewDelayedSnapshot:
        FTrace := TraceRecaptureAfterReset;
        FResetSubjects := FALSE;
        FInput[-2] := -100;
        FInput[-1] := 40;
        FInput[0] := 20;
        FInput[1] := 100;
        FExpectedImmediateFirst := 40;
        FExpectedImmediateSecond := 20;
        FExpectedDelayedFirst := 40;
        FExpectedDelayedSecond := 20;
        FImmediateEnable := TRUE;
        FImmediateResult := E_Result.Passed;
        FImmediateObservation := TRUE;
        FImmediateEvaluation := TRUE;
        FDelayedEnable := TRUE;
        FDelayedResult := E_Result.NotEvaluated;
        FDelayedObservation := TRUE;
        FDelayedEvaluation := FALSE;
    StepNewSnapshotMatches:
        FTrace := TraceRecaptureAfterReset;
        FResetSubjects := FALSE;
        FInput[-2] := -100;
        FInput[-1] := 40;
        FInput[0] := 20;
        FInput[1] := 100;
        FExpectedImmediateFirst := 40;
        FExpectedImmediateSecond := 20;
        FExpectedDelayedFirst := 40;
        FExpectedDelayedSecond := 20;
        FImmediateEnable := TRUE;
        FImmediateResult := E_Result.Passed;
        FImmediateObservation := TRUE;
        FImmediateEvaluation := TRUE;
        FDelayedEnable := TRUE;
        FDelayedResult := E_Result.Passed;
        FDelayedObservation := TRUE;
        FDelayedEvaluation := TRUE;
ELSE
    Error(Message := 'Unknown observation checkpoint.');
    RETURN;
END_CASE;
SelectStep := TRUE;
END_METHOD

END_FUNCTION_BLOCK

// ---- Framework/Assertions/POU/Arrays/DInt/AssertArrayNoValueChange_DInt.TcPOU
{region 'Documentation'}
(*!
<summary>Captures one snapshot until Reset; Disable/Re-Enable never replaces it.</summary>
<description>

Disabling observation preserves the original snapshot. Re-enabling requires a fresh
preceding observation before comparisons resume; it does not replace that snapshot.

StartIndex is an absolute IN index and Length selects 1..255 elements within IN. Memory
must have at least Length elements from its own lower bound. Invalid references or ranges
report Error.

The caller provides dedicated writable Memory that must not overlap IN; overlap is not
checked. Keep bindings, selected range and snapshot contents stable until Reset. Reset
invalidates the snapshot without clearing Memory bytes.

</description>
*)
{endregion}
FUNCTION_BLOCK AssertArrayNoValueChange_DInt EXTENDS AssertionBase
VAR_INPUT
    StartIndex : DINT; //! First selected index in IN; uses the array's declared index range, not a zero-based offset.
    Length : USINT; //! Number of monitored elements, from 1 through 255.
END_VAR
VAR_IN_OUT CONSTANT
    IN : ARRAY[*] OF DINT; //! Read-only actual data; the selected range must remain stable during the call.
END_VAR
VAR_IN_OUT
    Memory : ARRAY[*] OF DINT; //! Dedicated snapshot storage; only this assertion writes its selected elements.
END_VAR
VAR
    FSnapshotValid : BOOL;
    FObservationPrevious : BOOL;
    FEvaluationActive : BOOL;
END_VAR

SUPER^();

{region 'Documentation'}
(*!
<summary>Capture once or compare against the retained snapshot after range validation.</summary>
*)
{endregion}
METHOD PROTECTED Assert
VAR
    InLowerIndex : DINT;
    InUpperIndex : DINT;
    MemoryLowerIndex : DINT;
    MemoryUpperIndex : DINT;
    MemoryEndIndex : LINT;
    EndIndex : LINT;
    Offset : LINT;
    InIndex : DINT;
    MemoryIndex : DINT;
    Message : STRING(GVL_Constants.MessageLength);
    ReferenceText : STRING(GVL_Constants.AssertionValueLength);
    ActualText : STRING(GVL_Constants.AssertionValueLength);
END_VAR
FEvaluationActive := ObservationActive AND FObservationPrevious AND FSnapshotValid;
FObservationPrevious := ObservationActive;

IF NOT ObservationActive THEN
    RETURN;
END_IF;

IF Result = E_Result.Error THEN
    RETURN;
END_IF;

// C0371: FB inputs are checked here before any reference access.
{warning disable C0371}
IF NOT __ISVALIDREF(IN) THEN
    Error(Message := 'Assertion error: IN reference is invalid.');
    RETURN;
END_IF;

IF NOT __ISVALIDREF(Memory) THEN
    Error(Message := 'Assertion error: Memory reference is invalid.');
    RETURN;
END_IF;

InLowerIndex := LOWER_BOUND(IN, 1);
InUpperIndex := UPPER_BOUND(IN, 1);
MemoryLowerIndex := LOWER_BOUND(Memory, 1);
MemoryUpperIndex := UPPER_BOUND(Memory, 1);
EndIndex := DINT_TO_LINT(StartIndex) + USINT_TO_LINT(Length) - 1;
MemoryEndIndex := DINT_TO_LINT(MemoryLowerIndex) + USINT_TO_LINT(Length) - 1;

IF (Length = 0)
    OR (StartIndex < InLowerIndex) OR (StartIndex > InUpperIndex)
    OR (EndIndex > DINT_TO_LINT(InUpperIndex))
    OR (MemoryEndIndex > DINT_TO_LINT(MemoryUpperIndex)) THEN
    Message := CONCAT('Assertion error: array or memory range is invalid. StartIndex = ',
        DINT_TO_STRING(StartIndex));
    Message := CONCAT(Message, ', EndIndex = ');
    Message := CONCAT(Message, LINT_TO_STRING(EndIndex));
    Message := CONCAT(Message, ', Length = ');
    Message := CONCAT(Message, USINT_TO_STRING(Length));
    Message := CONCAT(Message, '.');
    Error(Message := Message);
    RETURN;
END_IF;

IF NOT FSnapshotValid THEN
    FOR Offset := 0 TO USINT_TO_LINT(Length) - 1 DO
        InIndex := LINT_TO_DINT(DINT_TO_LINT(StartIndex) + Offset);
        MemoryIndex := LINT_TO_DINT(DINT_TO_LINT(MemoryLowerIndex) + Offset);
        Memory[MemoryIndex] := IN[InIndex];
    END_FOR;
    FSnapshotValid := TRUE;
    RETURN;
END_IF;

IF NOT EvaluationActive THEN
    RETURN;
END_IF;

IF Result = E_Result.Failed THEN
    RETURN;
END_IF;

FOR Offset := 0 TO USINT_TO_LINT(Length) - 1 DO
    InIndex := LINT_TO_DINT(DINT_TO_LINT(StartIndex) + Offset);
    MemoryIndex := LINT_TO_DINT(DINT_TO_LINT(MemoryLowerIndex) + Offset);
    IF IN[InIndex] <> Memory[MemoryIndex] THEN
        ReferenceText := DINT_TO_STRING(Memory[MemoryIndex]);
        ActualText := DINT_TO_STRING(IN[InIndex]);
        Message := CONCAT('Assertion failed: array value changed. Reference[',
            DINT_TO_STRING(MemoryIndex));
        Message := CONCAT(Message, '] = ');
        Message := CONCAT(Message, ReferenceText);
        Message := CONCAT(Message, ', IN[');
        Message := CONCAT(Message, DINT_TO_STRING(InIndex));
        Message := CONCAT(Message, '] = ');
        Message := CONCAT(Message, ActualText);
        Message := CONCAT(Message, '.');
        Fail(Message := Message);
        RETURN;
    END_IF;
END_FOR;

Pass();
{warning restore C0371}
END_METHOD

{region 'Documentation'}
(*!
<summary>Current/last call has consecutive observation and an existing snapshot.</summary>
*)
{endregion}
{attribute 'monitoring' := 'call'}
PROPERTY PUBLIC EvaluationActive : BOOL //! Current/last call has consecutive observation and an existing snapshot.
GET // PUBLIC
EvaluationActive := FEvaluationActive;
END_GET
END_PROPERTY

{region 'Documentation'}
(*!
<summary>Invalidate the snapshot and observation history.</summary>
<description>

Does not clear external Memory. The next active observation captures a new snapshot
before comparison.

</description>
*)
{endregion}
METHOD PROTECTED ResetAssertion
FSnapshotValid := FALSE;
FObservationPrevious := FALSE;
FEvaluationActive := FALSE;
END_METHOD

END_FUNCTION_BLOCK

// ---- SelfTests/TestCases/TestSuite_AssertionObservation/Test_AssertionFloatingSnapshot.TcPOU
{region 'Documentation'}
(*!
<summary>Checks REAL/LREAL snapshot capture policy and comparison against the original values.</summary>
<description>
The second selected NaN must reject the complete capture without modifying even
the first Memory element. Signed infinities are valid array snapshots; later NaN
is a mismatch, not a capture error. Exactly representable tolerance steps separate
comparison against the original snapshot from comparison against the previous call.
IEEE union views only construct stimuli and inspect copied bits; no test arithmetic
or conversion is performed on non-finite values.
Each named step calls each subject once and checks public gates, result and local
findings before advancing in the next cycle. Outer Assertions collect checkpoints
per trace; subjects never contribute their intentional failures to the test result.
FirstFailedStep retains the first mismatch. No timed stimulus or expected-result
algorithm is used.
</description>
*)
{endregion}
FUNCTION_BLOCK Test_AssertionFloatingSnapshot EXTENDS TestCaseBase
VAR
    FReal : AssertArrayNoValueChange_Real;
    FLReal : AssertArrayNoValueChange_LReal;
    FRealInput : ARRAY[-1..0] OF REAL;
    FRealMemory : ARRAY[5..7] OF REAL;
    FRealFirst : AssertionRealRepresentation;
    FRealSecond : AssertionRealRepresentation;
    FRealMemoryFirst : AssertionRealRepresentation;
    FRealMemorySecond : AssertionRealRepresentation;
    FRealExpectedFirst : DWORD;
    FRealExpectedSecond : DWORD;
    FLRealInput : ARRAY[-1..0] OF LREAL;
    FLRealMemory : ARRAY[5..7] OF LREAL;
    FLRealFirst : AssertionLRealRepresentation;
    FLRealSecond : AssertionLRealRepresentation;
    FLRealMemoryFirst : AssertionLRealRepresentation;
    FLRealMemorySecond : AssertionLRealRepresentation;
    FLRealExpectedFirst : LWORD;
    FLRealExpectedSecond : LWORD;
    FCapture : EventBuffer;
    FEvents : ARRAY[1..CaptureLength] OF ST_Event;
    FCaptureFifo : ST_FifoStatus;
    FCaptureStatus : ST_EventBufferStatus;
    FSetupValid : BOOL;
    FStep : UINT;
    FTrace : UINT;
    FFirstFailedStep : UINT;
    FChecked : BOOL;
    FObservationReady : BOOL;
    FStepMatches : BOOL;
    FResultsMatch : BOOL;
    FActivityMatches : BOOL;
    FFindingsMatch : BOOL;
    FMemoryMatches : BOOL;
    FResetSubjects : BOOL;
    FRealEnable : BOOL;
    FRealResult : E_Result;
    FRealObservation : BOOL;
    FRealEvaluation : BOOL;
    FRealFinding : E_Result;
    FLRealEnable : BOOL;
    FLRealResult : E_Result;
    FLRealObservation : BOOL;
    FLRealEvaluation : BOOL;
    FLRealFinding : E_Result;
    FRejectedSnapshot : AssertTrue;
    FInfiniteSnapshot : AssertTrue;
    FLaterNaNDivergence : AssertTrue;
    FOriginalSnapshotTolerance : AssertTrue;
    FNewSnapshotAfterReset : AssertTrue;
END_VAR
VAR CONSTANT
    CaptureLength : UINT := 8;
    StepResetNaNCapture : UINT := 1;
    StepRejectNaNBeforeCopy : UINT := 2;
    StepNoRepeatedNaNEvent : UINT := 3;
    StepResetRejectedSnapshot : UINT := 4;
    StepRecoverCapture : UINT := 5;
    StepRecoverComparison : UINT := 6;
    StepResetInfinity : UINT := 7;
    StepCaptureInfinities : UINT := 8;
    StepEqualSignedInfinities : UINT := 9;
    StepChangedInfinitySign : UINT := 10;
    StepReturnToSignedInfinities : UINT := 11;
    StepResetLaterNaN : UINT := 12;
    StepCaptureBeforeLaterNaN : UINT := 13;
    StepCompareBeforeLaterNaN : UINT := 14;
    StepLaterNaNIsFailed : UINT := 15;
    StepResetTolerance : UINT := 16;
    StepCaptureTolerance : UINT := 17;
    StepWithinTolerance : UINT := 18;
    StepInclusiveTolerance : UINT := 19;
    StepBeyondOriginalTolerance : UINT := 20;
    StepResetNewFinite : UINT := 21;
    StepCaptureNewFinite : UINT := 22;
    StepCompareNewFinite : UINT := 23;
    LastStep : UINT := StepCompareNewFinite;
    TraceRejectedSnapshot : UINT := 1;
    TraceInfiniteSnapshot : UINT := 2;
    TraceLaterNaNDivergence : UINT := 3;
    TraceOriginalSnapshotTolerance : UINT := 4;
    TraceNewSnapshotAfterReset : UINT := 5;
END_VAR

SUPER^();

{region 'Documentation'}
(*!
<summary>Aggregates only the outer checks, not the intentionally failing subjects.</summary>
*)
{endregion}
METHOD PROTECTED AggregateResults
VAR_INPUT
    Aggregator : I_ResultAggregator; //! Borrowed result sink owned by the outer Test Case; add this test's checking Assertions without resetting or retaining the sink.
END_VAR
Aggregator.AddProvider(Provider := FRejectedSnapshot);
Aggregator.AddProvider(Provider := FInfiniteSnapshot);
Aggregator.AddProvider(Provider := FLaterNaNDivergence);
Aggregator.AddProvider(Provider := FOriginalSnapshotTolerance);
Aggregator.AddProvider(Provider := FNewSnapshotAfterReset);
END_METHOD

{region 'Documentation'}
(*!
<summary>Calls each production subject with stable bindings and the selected stimulus.</summary>
*)
{endregion}
METHOD PRIVATE CallSubjects
FReal(Enable := FRealEnable,
    State := E_State.Running,
    Tolerance := 0.5,
    StartIndex := -1,
    Length := 2,
    IN := FRealInput,
    Memory := FRealMemory);
FLReal(Enable := FLRealEnable,
    State := E_State.Running,
    Tolerance := 0.5,
    StartIndex := -1,
    Length := 2,
    IN := FLRealInput,
    Memory := FLRealMemory);
END_METHOD

{region 'Documentation'}
(*!
<summary>Checks finding order, identities and exact count without retaining prior events.</summary>
*)
{endregion}
METHOD PRIVATE CheckFindings
VAR
    Index : UINT;
    FindingMatches : BOOL;
END_VAR
Index := 1;
FFindingsMatch := TRUE;
IF FRealFinding <> E_Result.NotEvaluated THEN
    FindingMatches := IsFindingValid(Index := Index,
        ExpectedName := FReal.Name,
        ExpectedResult := FRealFinding);
    FFindingsMatch := FFindingsMatch AND FindingMatches;
    Index := Index + 1;
END_IF;
IF FLRealFinding <> E_Result.NotEvaluated THEN
    FindingMatches := IsFindingValid(Index := Index,
        ExpectedName := FLReal.Name,
        ExpectedResult := FLRealFinding);
    FFindingsMatch := FFindingsMatch AND FindingMatches;
    Index := Index + 1;
END_IF;
FFindingsMatch := FFindingsMatch
    AND (FCaptureStatus.SequenceId = UINT_TO_UDINT(Index - 1))
    AND (FCaptureStatus.LostEventCount = 0);
END_METHOD

{region 'Documentation'}
(*!
<summary>Rejects an incomplete capture or subject setup.</summary>
*)
{endregion}
METHOD PROTECTED CheckInitialization : BOOL //! TRUE when the inherited initialization check and this concrete fixture check both accept the setup.
CheckInitialization := SUPER^.CheckInitialization();
IF NOT CheckInitialization THEN
    RETURN;
END_IF;

CheckInitialization := FSetupValid
    AND FRejectedSnapshot.IsInitialized
    AND FInfiniteSnapshot.IsInitialized
    AND FLaterNaNDivergence.IsInitialized
    AND FOriginalSnapshotTolerance.IsInitialized
    AND FNewSnapshotAfterReset.IsInitialized;
IF NOT CheckInitialization THEN
    EventPublisher.PublishEvent(Event := CreateFrameworkEvent(Name := Name,
        ResourceName := '',
        State := State,
        Severity := E_EventSeverity.Error,
        Message := 'Observation selftest setup failed.'));
END_IF;
END_METHOD

{region 'Documentation'}
(*!
<summary>Checks copied IEEE representations without evaluating non-finite floating-point values.</summary>
*)
{endregion}
METHOD PRIVATE CheckMemory
FRealMemoryFirst.Value := FRealMemory[5];
FRealMemorySecond.Value := FRealMemory[6];
FLRealMemoryFirst.Value := FLRealMemory[5];
FLRealMemorySecond.Value := FLRealMemory[6];
FMemoryMatches := (FRealMemoryFirst.Bits = FRealExpectedFirst)
    AND (FRealMemorySecond.Bits = FRealExpectedSecond)
    AND (FRealMemory[7] = -999.0)
    AND (FLRealMemoryFirst.Bits = FLRealExpectedFirst)
    AND (FLRealMemorySecond.Bits = FLRealExpectedSecond)
    AND (FLRealMemory[7] = -999.0);
END_METHOD

{region 'Documentation'}
(*!
<summary>Checks literal result and observation/evaluation expectations.</summary>
*)
{endregion}
METHOD PRIVATE CheckResults
FResultsMatch := (FReal.Result = FRealResult)
    AND (FLReal.Result = FLRealResult);
FActivityMatches := (FReal.Enabled = FRealEnable)
    AND (FReal.ObservationActive = FRealObservation)
    AND (FReal.EvaluationActive = FRealEvaluation)
    AND (FLReal.Enabled = FLRealEnable)
    AND (FLReal.ObservationActive = FLRealObservation)
    AND (FLReal.EvaluationActive = FLRealEvaluation);
END_METHOD

{region 'Documentation'}
(*!
<summary>Initializes outer checks and isolates intentional subject findings.</summary>
*)
{endregion}
METHOD PROTECTED Configure
VAR
    Initialized : BOOL;
END_VAR
FPreparationStateCount := 0;
FTestStateCount := 1;
FRejectedSnapshot.Initialize(Parent := THIS^,
    AssertionName := 'RejectedSnapshot');
FInfiniteSnapshot.Initialize(Parent := THIS^,
    AssertionName := 'InfiniteSnapshot');
FLaterNaNDivergence.Initialize(Parent := THIS^,
    AssertionName := 'LaterNaNDivergence');
FOriginalSnapshotTolerance.Initialize(Parent := THIS^,
    AssertionName := 'OriginalSnapshotTolerance');
FNewSnapshotAfterReset.Initialize(Parent := THIS^,
    AssertionName := 'NewSnapshotAfterReset');
FSetupValid := FCapture.Initialize(Buffer := FEvents,
    FifoControl := FCaptureFifo,
    Status := FCaptureStatus);
FReal.BindPublisher(Publisher := FCapture);
Initialized := FReal.Initialize(Parent := THIS^,
    AssertionName := 'Real',
    ObserveFirstCycle := TRUE);
FSetupValid := FSetupValid AND Initialized;
FLReal.BindPublisher(Publisher := FCapture);
Initialized := FLReal.Initialize(Parent := THIS^,
    AssertionName := 'LReal',
    ObserveFirstCycle := TRUE);
FSetupValid := FSetupValid AND Initialized;
END_METHOD

{region 'Documentation'}
(*!
<summary>Checks one expected Failed or Error finding from the bounded local capture.</summary>
*)
{endregion}
METHOD PRIVATE IsFindingValid : BOOL //! TRUE when the selected captured finding satisfies the scenario metadata and diagnostic checks.
VAR_INPUT
    Index : UINT; //! One-based index in the retained isolated event capture.
    ExpectedName : STRING(GVL_Constants.NameLength); //! Independently authored Assertion name expected in the selected finding.
    ExpectedResult : E_Result; //! Independently authored finding result.
END_VAR
IsFindingValid := (FEvents[Index].SequenceId = UINT_TO_UDINT(Index))
    AND (FEvents[Index].Name = ExpectedName)
    AND (FEvents[Index].OwnerScope = E_OwnerScope.Assertion)
    AND (FEvents[Index].EventType = E_EventType.Result)
    AND (FEvents[Index].State = E_State.Running)
    AND (FEvents[Index].Result = ExpectedResult)
    AND (FEvents[Index].Message <> '');
END_METHOD

{region 'Documentation'}
(*!
<summary>Completes abort without asynchronous resources.</summary>
*)
{endregion}
METHOD PROTECTED ProcessAbort
VAR_INPUT
    Enable : BOOL; //! Phase permission supplied by the owning Test Case; FALSE does not authorize progression, while observation may continue.
END_VAR
IF Enable THEN
    CompleteAbort();
END_IF;
END_METHOD

{region 'Documentation'}
(*!
<summary>Checks this checkpoint before the next cycle advances the trace.</summary>
*)
{endregion}
METHOD PROTECTED ProcessAssertions
VAR_INPUT
    Enable : BOOL; //! Phase permission supplied by the owning Test Case; FALSE does not authorize progression, while observation may continue.
END_VAR
VAR
    Check : BOOL;
END_VAR
Check := Enable AND FObservationReady;
FRejectedSnapshot(Enable := Check AND (FTrace = TraceRejectedSnapshot),
    State := State,
    IN := FStepMatches);
FInfiniteSnapshot(Enable := Check AND (FTrace = TraceInfiniteSnapshot),
    State := State,
    IN := FStepMatches);
FLaterNaNDivergence(Enable := Check AND (FTrace = TraceLaterNaNDivergence),
    State := State,
    IN := FStepMatches);
FOriginalSnapshotTolerance(Enable := Check AND (FTrace = TraceOriginalSnapshotTolerance),
    State := State,
    IN := FStepMatches);
FNewSnapshotAfterReset(Enable := Check AND (FTrace = TraceNewSnapshotAfterReset),
    State := State,
    IN := FStepMatches);
IF Check THEN
    FChecked := TRUE;
END_IF;
END_METHOD

{region 'Documentation'}
(*!
<summary>No Preparation phase is required.</summary>
*)
{endregion}
METHOD PROTECTED ProcessPreparations
VAR_INPUT
    // SA0033: Required hook; this test has no Preparation phase.
    {attribute 'analysis' := '-33'}
    Enable : BOOL; //! Phase permission supplied by the owning Test Case; FALSE does not authorize progression, while observation may continue.
END_VAR
END_METHOD

{region 'Documentation'}
(*!
<summary>Resets checkpoint bookkeeping and queues each subject reset.</summary>
*)
{endregion}
METHOD PROTECTED ProcessReset
FStep := StepResetNaNCapture;
FTrace := 0;
FFirstFailedStep := 0;
FChecked := FALSE;
FObservationReady := FALSE;
FCapture.Reset();
ResetSubjects();
FRejectedSnapshot.Reset();
FInfiniteSnapshot.Reset();
FLaterNaNDivergence.Reset();
FOriginalSnapshotTolerance.Reset();
FNewSnapshotAfterReset.Reset();
CompleteReset();
END_METHOD

{region 'Documentation'}
(*!
<summary>Executes exactly one named checkpoint per active PLC cycle.</summary>
*)
{endregion}
METHOD PROTECTED ProcessTests
VAR_INPUT
    Enable : BOOL; //! Phase permission supplied by the owning Test Case; FALSE does not authorize progression, while observation may continue.
END_VAR
IF NOT Enable THEN
    RETURN;
END_IF;

IF FChecked THEN
    FChecked := FALSE;
    FObservationReady := FALSE;
    IF FStep = LastStep THEN
        CompleteTests();
        RETURN;
    END_IF;
    FStep := FStep + 1;
END_IF;

IF NOT SelectStep() THEN
    RETURN;
END_IF;
FCapture.Reset();
IF FResetSubjects THEN
    ResetSubjects();
END_IF;
CallSubjects();
CheckResults();
CheckMemory();
CheckFindings();
FStepMatches := FResultsMatch AND FActivityMatches AND FMemoryMatches AND FFindingsMatch;
IF NOT FStepMatches AND (FFirstFailedStep = 0) THEN
    FFirstFailedStep := FStep;
END_IF;
FObservationReady := TRUE;
END_METHOD

{region 'Documentation'}
(*!
<summary>Queues subject reset; the next bound call consumes it.</summary>
*)
{endregion}
METHOD PRIVATE ResetSubjects
FReal.Reset();
FLReal.Reset();
END_METHOD

{region 'Documentation'}
(*!
<summary>Selects literal stimuli, gates and findings for a named checkpoint.</summary>
*)
{endregion}
METHOD PRIVATE SelectStep : BOOL //! TRUE after selecting a supported script step and its literal expectations; FALSE reports an unknown step.
SelectStep := FALSE;
FRealFinding := E_Result.NotEvaluated;
FLRealFinding := E_Result.NotEvaluated;
CASE FStep OF
    StepResetNaNCapture:
        FTrace := TraceRejectedSnapshot;
        FResetSubjects := TRUE;
        FRealFirst.Bits := DWORD#16#41000000;
        FRealSecond.Bits := DWORD#16#7FC00000;
        FRealInput[-1] := FRealFirst.Value;
        FRealInput[0] := FRealSecond.Value;
        FRealExpectedFirst := DWORD#16#C4424000;
        FRealExpectedSecond := DWORD#16#C45E0000;
        FRealMemory[5] := -777.0;
        FRealMemory[6] := -888.0;
        FRealMemory[7] := -999.0;
        FLRealFirst.Bits := LWORD#16#4020000000000000;
        FLRealSecond.Bits := LWORD#16#7FF8000000000000;
        FLRealInput[-1] := FLRealFirst.Value;
        FLRealInput[0] := FLRealSecond.Value;
        FLRealExpectedFirst := LWORD#16#C088480000000000;
        FLRealExpectedSecond := LWORD#16#C08BC00000000000;
        FLRealMemory[5] := -777.0;
        FLRealMemory[6] := -888.0;
        FLRealMemory[7] := -999.0;
        FRealEnable := TRUE;
        FRealResult := E_Result.NotEvaluated;
        FRealObservation := FALSE;
        FRealEvaluation := FALSE;
        FLRealEnable := TRUE;
        FLRealResult := E_Result.NotEvaluated;
        FLRealObservation := FALSE;
        FLRealEvaluation := FALSE;
    StepRejectNaNBeforeCopy:
        FTrace := TraceRejectedSnapshot;
        FResetSubjects := FALSE;
        FRealFirst.Bits := DWORD#16#41000000;
        FRealSecond.Bits := DWORD#16#7FC00000;
        FRealInput[-1] := FRealFirst.Value;
        FRealInput[0] := FRealSecond.Value;
        FRealExpectedFirst := DWORD#16#C4424000;
        FRealExpectedSecond := DWORD#16#C45E0000;
        FLRealFirst.Bits := LWORD#16#4020000000000000;
        FLRealSecond.Bits := LWORD#16#7FF8000000000000;
        FLRealInput[-1] := FLRealFirst.Value;
        FLRealInput[0] := FLRealSecond.Value;
        FLRealExpectedFirst := LWORD#16#C088480000000000;
        FLRealExpectedSecond := LWORD#16#C08BC00000000000;
        FRealEnable := TRUE;
        FRealResult := E_Result.Error;
        FRealObservation := TRUE;
        FRealEvaluation := FALSE;
        FRealFinding := E_Result.Error;
        FLRealEnable := TRUE;
        FLRealResult := E_Result.Error;
        FLRealObservation := TRUE;
        FLRealEvaluation := FALSE;
        FLRealFinding := E_Result.Error;
    StepNoRepeatedNaNEvent:
        FTrace := TraceRejectedSnapshot;
        FResetSubjects := FALSE;
        FRealFirst.Bits := DWORD#16#41000000;
        FRealSecond.Bits := DWORD#16#7FC00000;
        FRealInput[-1] := FRealFirst.Value;
        FRealInput[0] := FRealSecond.Value;
        FRealExpectedFirst := DWORD#16#C4424000;
        FRealExpectedSecond := DWORD#16#C45E0000;
        FLRealFirst.Bits := LWORD#16#4020000000000000;
        FLRealSecond.Bits := LWORD#16#7FF8000000000000;
        FLRealInput[-1] := FLRealFirst.Value;
        FLRealInput[0] := FLRealSecond.Value;
        FLRealExpectedFirst := LWORD#16#C088480000000000;
        FLRealExpectedSecond := LWORD#16#C08BC00000000000;
        FRealEnable := TRUE;
        FRealResult := E_Result.Error;
        FRealObservation := TRUE;
        FRealEvaluation := FALSE;
        FLRealEnable := TRUE;
        FLRealResult := E_Result.Error;
        FLRealObservation := TRUE;
        FLRealEvaluation := FALSE;
    StepResetRejectedSnapshot:
        FTrace := TraceRejectedSnapshot;
        FResetSubjects := TRUE;
        FRealFirst.Bits := DWORD#16#41000000;
        FRealSecond.Bits := DWORD#16#41A00000;
        FRealInput[-1] := FRealFirst.Value;
        FRealInput[0] := FRealSecond.Value;
        FRealExpectedFirst := DWORD#16#C4424000;
        FRealExpectedSecond := DWORD#16#C45E0000;
        FLRealFirst.Bits := LWORD#16#4020000000000000;
        FLRealSecond.Bits := LWORD#16#4034000000000000;
        FLRealInput[-1] := FLRealFirst.Value;
        FLRealInput[0] := FLRealSecond.Value;
        FLRealExpectedFirst := LWORD#16#C088480000000000;
        FLRealExpectedSecond := LWORD#16#C08BC00000000000;
        FRealEnable := TRUE;
        FRealResult := E_Result.NotEvaluated;
        FRealObservation := FALSE;
        FRealEvaluation := FALSE;
        FLRealEnable := TRUE;
        FLRealResult := E_Result.NotEvaluated;
        FLRealObservation := FALSE;
        FLRealEvaluation := FALSE;
    StepRecoverCapture:
        FTrace := TraceRejectedSnapshot;
        FResetSubjects := FALSE;
        FRealFirst.Bits := DWORD#16#41000000;
        FRealSecond.Bits := DWORD#16#41A00000;
        FRealInput[-1] := FRealFirst.Value;
        FRealInput[0] := FRealSecond.Value;
        FRealExpectedFirst := DWORD#16#41000000;
        FRealExpectedSecond := DWORD#16#41A00000;
        FLRealFirst.Bits := LWORD#16#4020000000000000;
        FLRealSecond.Bits := LWORD#16#4034000000000000;
        FLRealInput[-1] := FLRealFirst.Value;
        FLRealInput[0] := FLRealSecond.Value;
        FLRealExpectedFirst := LWORD#16#4020000000000000;
        FLRealExpectedSecond := LWORD#16#4034000000000000;
        FRealEnable := TRUE;
        FRealResult := E_Result.NotEvaluated;
        FRealObservation := TRUE;
        FRealEvaluation := FALSE;
        FLRealEnable := TRUE;
        FLRealResult := E_Result.NotEvaluated;
        FLRealObservation := TRUE;
        FLRealEvaluation := FALSE;
    StepRecoverComparison:
        FTrace := TraceRejectedSnapshot;
        FResetSubjects := FALSE;
        FRealFirst.Bits := DWORD#16#41000000;
        FRealSecond.Bits := DWORD#16#41A00000;
        FRealInput[-1] := FRealFirst.Value;
        FRealInput[0] := FRealSecond.Value;
        FRealExpectedFirst := DWORD#16#41000000;
        FRealExpectedSecond := DWORD#16#41A00000;
        FLRealFirst.Bits := LWORD#16#4020000000000000;
        FLRealSecond.Bits := LWORD#16#4034000000000000;
        FLRealInput[-1] := FLRealFirst.Value;
        FLRealInput[0] := FLRealSecond.Value;
        FLRealExpectedFirst := LWORD#16#4020000000000000;
        FLRealExpectedSecond := LWORD#16#4034000000000000;
        FRealEnable := TRUE;
        FRealResult := E_Result.Passed;
        FRealObservation := TRUE;
        FRealEvaluation := TRUE;
        FLRealEnable := TRUE;
        FLRealResult := E_Result.Passed;
        FLRealObservation := TRUE;
        FLRealEvaluation := TRUE;
    StepResetInfinity:
        FTrace := TraceInfiniteSnapshot;
        FResetSubjects := TRUE;
        FRealFirst.Bits := DWORD#16#7F800000;
        FRealSecond.Bits := DWORD#16#FF800000;
        FRealInput[-1] := FRealFirst.Value;
        FRealInput[0] := FRealSecond.Value;
        FRealExpectedFirst := DWORD#16#41000000;
        FRealExpectedSecond := DWORD#16#41A00000;
        FLRealFirst.Bits := LWORD#16#7FF0000000000000;
        FLRealSecond.Bits := LWORD#16#FFF0000000000000;
        FLRealInput[-1] := FLRealFirst.Value;
        FLRealInput[0] := FLRealSecond.Value;
        FLRealExpectedFirst := LWORD#16#4020000000000000;
        FLRealExpectedSecond := LWORD#16#4034000000000000;
        FRealEnable := TRUE;
        FRealResult := E_Result.NotEvaluated;
        FRealObservation := FALSE;
        FRealEvaluation := FALSE;
        FLRealEnable := TRUE;
        FLRealResult := E_Result.NotEvaluated;
        FLRealObservation := FALSE;
        FLRealEvaluation := FALSE;
    StepCaptureInfinities:
        FTrace := TraceInfiniteSnapshot;
        FResetSubjects := FALSE;
        FRealFirst.Bits := DWORD#16#7F800000;
        FRealSecond.Bits := DWORD#16#FF800000;
        FRealInput[-1] := FRealFirst.Value;
        FRealInput[0] := FRealSecond.Value;
        FRealExpectedFirst := DWORD#16#7F800000;
        FRealExpectedSecond := DWORD#16#FF800000;
        FLRealFirst.Bits := LWORD#16#7FF0000000000000;
        FLRealSecond.Bits := LWORD#16#FFF0000000000000;
        FLRealInput[-1] := FLRealFirst.Value;
        FLRealInput[0] := FLRealSecond.Value;
        FLRealExpectedFirst := LWORD#16#7FF0000000000000;
        FLRealExpectedSecond := LWORD#16#FFF0000000000000;
        FRealEnable := TRUE;
        FRealResult := E_Result.NotEvaluated;
        FRealObservation := TRUE;
        FRealEvaluation := FALSE;
        FLRealEnable := TRUE;
        FLRealResult := E_Result.NotEvaluated;
        FLRealObservation := TRUE;
        FLRealEvaluation := FALSE;
    StepEqualSignedInfinities:
        FTrace := TraceInfiniteSnapshot;
        FResetSubjects := FALSE;
        FRealFirst.Bits := DWORD#16#7F800000;
        FRealSecond.Bits := DWORD#16#FF800000;
        FRealInput[-1] := FRealFirst.Value;
        FRealInput[0] := FRealSecond.Value;
        FRealExpectedFirst := DWORD#16#7F800000;
        FRealExpectedSecond := DWORD#16#FF800000;
        FLRealFirst.Bits := LWORD#16#7FF0000000000000;
        FLRealSecond.Bits := LWORD#16#FFF0000000000000;
        FLRealInput[-1] := FLRealFirst.Value;
        FLRealInput[0] := FLRealSecond.Value;
        FLRealExpectedFirst := LWORD#16#7FF0000000000000;
        FLRealExpectedSecond := LWORD#16#FFF0000000000000;
        FRealEnable := TRUE;
        FRealResult := E_Result.Passed;
        FRealObservation := TRUE;
        FRealEvaluation := TRUE;
        FLRealEnable := TRUE;
        FLRealResult := E_Result.Passed;
        FLRealObservation := TRUE;
        FLRealEvaluation := TRUE;
    StepChangedInfinitySign:
        FTrace := TraceInfiniteSnapshot;
        FResetSubjects := FALSE;
        FRealFirst.Bits := DWORD#16#7F800000;
        FRealSecond.Bits := DWORD#16#7F800000;
        FRealInput[-1] := FRealFirst.Value;
        FRealInput[0] := FRealSecond.Value;
        FRealExpectedFirst := DWORD#16#7F800000;
        FRealExpectedSecond := DWORD#16#FF800000;
        FLRealFirst.Bits := LWORD#16#7FF0000000000000;
        FLRealSecond.Bits := LWORD#16#7FF0000000000000;
        FLRealInput[-1] := FLRealFirst.Value;
        FLRealInput[0] := FLRealSecond.Value;
        FLRealExpectedFirst := LWORD#16#7FF0000000000000;
        FLRealExpectedSecond := LWORD#16#FFF0000000000000;
        FRealEnable := TRUE;
        FRealResult := E_Result.Failed;
        FRealObservation := TRUE;
        FRealEvaluation := TRUE;
        FRealFinding := E_Result.Failed;
        FLRealEnable := TRUE;
        FLRealResult := E_Result.Failed;
        FLRealObservation := TRUE;
        FLRealEvaluation := TRUE;
        FLRealFinding := E_Result.Failed;
    StepReturnToSignedInfinities:
        FTrace := TraceInfiniteSnapshot;
        FResetSubjects := FALSE;
        FRealFirst.Bits := DWORD#16#7F800000;
        FRealSecond.Bits := DWORD#16#FF800000;
        FRealInput[-1] := FRealFirst.Value;
        FRealInput[0] := FRealSecond.Value;
        FRealExpectedFirst := DWORD#16#7F800000;
        FRealExpectedSecond := DWORD#16#FF800000;
        FLRealFirst.Bits := LWORD#16#7FF0000000000000;
        FLRealSecond.Bits := LWORD#16#FFF0000000000000;
        FLRealInput[-1] := FLRealFirst.Value;
        FLRealInput[0] := FLRealSecond.Value;
        FLRealExpectedFirst := LWORD#16#7FF0000000000000;
        FLRealExpectedSecond := LWORD#16#FFF0000000000000;
        FRealEnable := TRUE;
        FRealResult := E_Result.Failed;
        FRealObservation := TRUE;
        FRealEvaluation := TRUE;
        FLRealEnable := TRUE;
        FLRealResult := E_Result.Failed;
        FLRealObservation := TRUE;
        FLRealEvaluation := TRUE;
    StepResetLaterNaN:
        FTrace := TraceLaterNaNDivergence;
        FResetSubjects := TRUE;
        FRealFirst.Bits := DWORD#16#41000000;
        FRealSecond.Bits := DWORD#16#41A00000;
        FRealInput[-1] := FRealFirst.Value;
        FRealInput[0] := FRealSecond.Value;
        FRealExpectedFirst := DWORD#16#7F800000;
        FRealExpectedSecond := DWORD#16#FF800000;
        FLRealFirst.Bits := LWORD#16#4020000000000000;
        FLRealSecond.Bits := LWORD#16#4034000000000000;
        FLRealInput[-1] := FLRealFirst.Value;
        FLRealInput[0] := FLRealSecond.Value;
        FLRealExpectedFirst := LWORD#16#7FF0000000000000;
        FLRealExpectedSecond := LWORD#16#FFF0000000000000;
        FRealEnable := TRUE;
        FRealResult := E_Result.NotEvaluated;
        FRealObservation := FALSE;
        FRealEvaluation := FALSE;
        FLRealEnable := TRUE;
        FLRealResult := E_Result.NotEvaluated;
        FLRealObservation := FALSE;
        FLRealEvaluation := FALSE;
    StepCaptureBeforeLaterNaN:
        FTrace := TraceLaterNaNDivergence;
        FResetSubjects := FALSE;
        FRealFirst.Bits := DWORD#16#41000000;
        FRealSecond.Bits := DWORD#16#41A00000;
        FRealInput[-1] := FRealFirst.Value;
        FRealInput[0] := FRealSecond.Value;
        FRealExpectedFirst := DWORD#16#41000000;
        FRealExpectedSecond := DWORD#16#41A00000;
        FLRealFirst.Bits := LWORD#16#4020000000000000;
        FLRealSecond.Bits := LWORD#16#4034000000000000;
        FLRealInput[-1] := FLRealFirst.Value;
        FLRealInput[0] := FLRealSecond.Value;
        FLRealExpectedFirst := LWORD#16#4020000000000000;
        FLRealExpectedSecond := LWORD#16#4034000000000000;
        FRealEnable := TRUE;
        FRealResult := E_Result.NotEvaluated;
        FRealObservation := TRUE;
        FRealEvaluation := FALSE;
        FLRealEnable := TRUE;
        FLRealResult := E_Result.NotEvaluated;
        FLRealObservation := TRUE;
        FLRealEvaluation := FALSE;
    StepCompareBeforeLaterNaN:
        FTrace := TraceLaterNaNDivergence;
        FResetSubjects := FALSE;
        FRealFirst.Bits := DWORD#16#41000000;
        FRealSecond.Bits := DWORD#16#41A00000;
        FRealInput[-1] := FRealFirst.Value;
        FRealInput[0] := FRealSecond.Value;
        FRealExpectedFirst := DWORD#16#41000000;
        FRealExpectedSecond := DWORD#16#41A00000;
        FLRealFirst.Bits := LWORD#16#4020000000000000;
        FLRealSecond.Bits := LWORD#16#4034000000000000;
        FLRealInput[-1] := FLRealFirst.Value;
        FLRealInput[0] := FLRealSecond.Value;
        FLRealExpectedFirst := LWORD#16#4020000000000000;
        FLRealExpectedSecond := LWORD#16#4034000000000000;
        FRealEnable := TRUE;
        FRealResult := E_Result.Passed;
        FRealObservation := TRUE;
        FRealEvaluation := TRUE;
        FLRealEnable := TRUE;
        FLRealResult := E_Result.Passed;
        FLRealObservation := TRUE;
        FLRealEvaluation := TRUE;
    StepLaterNaNIsFailed:
        FTrace := TraceLaterNaNDivergence;
        FResetSubjects := FALSE;
        FRealFirst.Bits := DWORD#16#41000000;
        FRealSecond.Bits := DWORD#16#7FC00000;
        FRealInput[-1] := FRealFirst.Value;
        FRealInput[0] := FRealSecond.Value;
        FRealExpectedFirst := DWORD#16#41000000;
        FRealExpectedSecond := DWORD#16#41A00000;
        FLRealFirst.Bits := LWORD#16#4020000000000000;
        FLRealSecond.Bits := LWORD#16#7FF8000000000000;
        FLRealInput[-1] := FLRealFirst.Value;
        FLRealInput[0] := FLRealSecond.Value;
        FLRealExpectedFirst := LWORD#16#4020000000000000;
        FLRealExpectedSecond := LWORD#16#4034000000000000;
        FRealEnable := TRUE;
        FRealResult := E_Result.Failed;
        FRealObservation := TRUE;
        FRealEvaluation := TRUE;
        FRealFinding := E_Result.Failed;
        FLRealEnable := TRUE;
        FLRealResult := E_Result.Failed;
        FLRealObservation := TRUE;
        FLRealEvaluation := TRUE;
        FLRealFinding := E_Result.Failed;
    StepResetTolerance:
        FTrace := TraceOriginalSnapshotTolerance;
        FResetSubjects := TRUE;
        FRealFirst.Bits := DWORD#16#41000000;
        FRealSecond.Bits := DWORD#16#41A00000;
        FRealInput[-1] := FRealFirst.Value;
        FRealInput[0] := FRealSecond.Value;
        FRealExpectedFirst := DWORD#16#41000000;
        FRealExpectedSecond := DWORD#16#41A00000;
        FLRealFirst.Bits := LWORD#16#4020000000000000;
        FLRealSecond.Bits := LWORD#16#4034000000000000;
        FLRealInput[-1] := FLRealFirst.Value;
        FLRealInput[0] := FLRealSecond.Value;
        FLRealExpectedFirst := LWORD#16#4020000000000000;
        FLRealExpectedSecond := LWORD#16#4034000000000000;
        FRealEnable := TRUE;
        FRealResult := E_Result.NotEvaluated;
        FRealObservation := FALSE;
        FRealEvaluation := FALSE;
        FLRealEnable := TRUE;
        FLRealResult := E_Result.NotEvaluated;
        FLRealObservation := FALSE;
        FLRealEvaluation := FALSE;
    StepCaptureTolerance:
        FTrace := TraceOriginalSnapshotTolerance;
        FResetSubjects := FALSE;
        FRealFirst.Bits := DWORD#16#41000000;
        FRealSecond.Bits := DWORD#16#41A00000;
        FRealInput[-1] := FRealFirst.Value;
        FRealInput[0] := FRealSecond.Value;
        FRealExpectedFirst := DWORD#16#41000000;
        FRealExpectedSecond := DWORD#16#41A00000;
        FLRealFirst.Bits := LWORD#16#4020000000000000;
        FLRealSecond.Bits := LWORD#16#4034000000000000;
        FLRealInput[-1] := FLRealFirst.Value;
        FLRealInput[0] := FLRealSecond.Value;
        FLRealExpectedFirst := LWORD#16#4020000000000000;
        FLRealExpectedSecond := LWORD#16#4034000000000000;
        FRealEnable := TRUE;
        FRealResult := E_Result.NotEvaluated;
        FRealObservation := TRUE;
        FRealEvaluation := FALSE;
        FLRealEnable := TRUE;
        FLRealResult := E_Result.NotEvaluated;
        FLRealObservation := TRUE;
        FLRealEvaluation := FALSE;
    StepWithinTolerance:
        FTrace := TraceOriginalSnapshotTolerance;
        FResetSubjects := FALSE;
        FRealFirst.Bits := DWORD#16#41040000;
        FRealSecond.Bits := DWORD#16#41A00000;
        FRealInput[-1] := FRealFirst.Value;
        FRealInput[0] := FRealSecond.Value;
        FRealExpectedFirst := DWORD#16#41000000;
        FRealExpectedSecond := DWORD#16#41A00000;
        FLRealFirst.Bits := LWORD#16#4020800000000000;
        FLRealSecond.Bits := LWORD#16#4034000000000000;
        FLRealInput[-1] := FLRealFirst.Value;
        FLRealInput[0] := FLRealSecond.Value;
        FLRealExpectedFirst := LWORD#16#4020000000000000;
        FLRealExpectedSecond := LWORD#16#4034000000000000;
        FRealEnable := TRUE;
        FRealResult := E_Result.Passed;
        FRealObservation := TRUE;
        FRealEvaluation := TRUE;
        FLRealEnable := TRUE;
        FLRealResult := E_Result.Passed;
        FLRealObservation := TRUE;
        FLRealEvaluation := TRUE;
    StepInclusiveTolerance:
        FTrace := TraceOriginalSnapshotTolerance;
        FResetSubjects := FALSE;
        FRealFirst.Bits := DWORD#16#41080000;
        FRealSecond.Bits := DWORD#16#41A00000;
        FRealInput[-1] := FRealFirst.Value;
        FRealInput[0] := FRealSecond.Value;
        FRealExpectedFirst := DWORD#16#41000000;
        FRealExpectedSecond := DWORD#16#41A00000;
        FLRealFirst.Bits := LWORD#16#4021000000000000;
        FLRealSecond.Bits := LWORD#16#4034000000000000;
        FLRealInput[-1] := FLRealFirst.Value;
        FLRealInput[0] := FLRealSecond.Value;
        FLRealExpectedFirst := LWORD#16#4020000000000000;
        FLRealExpectedSecond := LWORD#16#4034000000000000;
        FRealEnable := TRUE;
        FRealResult := E_Result.Passed;
        FRealObservation := TRUE;
        FRealEvaluation := TRUE;
        FLRealEnable := TRUE;
        FLRealResult := E_Result.Passed;
        FLRealObservation := TRUE;
        FLRealEvaluation := TRUE;
    StepBeyondOriginalTolerance:
        FTrace := TraceOriginalSnapshotTolerance;
        FResetSubjects := FALSE;
        FRealFirst.Bits := DWORD#16#410C0000;
        FRealSecond.Bits := DWORD#16#41A00000;
        FRealInput[-1] := FRealFirst.Value;
        FRealInput[0] := FRealSecond.Value;
        FRealExpectedFirst := DWORD#16#41000000;
        FRealExpectedSecond := DWORD#16#41A00000;
        FLRealFirst.Bits := LWORD#16#4021800000000000;
        FLRealSecond.Bits := LWORD#16#4034000000000000;
        FLRealInput[-1] := FLRealFirst.Value;
        FLRealInput[0] := FLRealSecond.Value;
        FLRealExpectedFirst := LWORD#16#4020000000000000;
        FLRealExpectedSecond := LWORD#16#4034000000000000;
        FRealEnable := TRUE;
        FRealResult := E_Result.Failed;
        FRealObservation := TRUE;
        FRealEvaluation := TRUE;
        FRealFinding := E_Result.Failed;
        FLRealEnable := TRUE;
        FLRealResult := E_Result.Failed;
        FLRealObservation := TRUE;
        FLRealEvaluation := TRUE;
        FLRealFinding := E_Result.Failed;
    StepResetNewFinite:
        FTrace := TraceNewSnapshotAfterReset;
        FResetSubjects := TRUE;
        FRealFirst.Bits := DWORD#16#42200000;
        FRealSecond.Bits := DWORD#16#42480000;
        FRealInput[-1] := FRealFirst.Value;
        FRealInput[0] := FRealSecond.Value;
        FRealExpectedFirst := DWORD#16#41000000;
        FRealExpectedSecond := DWORD#16#41A00000;
        FLRealFirst.Bits := LWORD#16#4044000000000000;
        FLRealSecond.Bits := LWORD#16#4049000000000000;
        FLRealInput[-1] := FLRealFirst.Value;
        FLRealInput[0] := FLRealSecond.Value;
        FLRealExpectedFirst := LWORD#16#4020000000000000;
        FLRealExpectedSecond := LWORD#16#4034000000000000;
        FRealEnable := TRUE;
        FRealResult := E_Result.NotEvaluated;
        FRealObservation := FALSE;
        FRealEvaluation := FALSE;
        FLRealEnable := TRUE;
        FLRealResult := E_Result.NotEvaluated;
        FLRealObservation := FALSE;
        FLRealEvaluation := FALSE;
    StepCaptureNewFinite:
        FTrace := TraceNewSnapshotAfterReset;
        FResetSubjects := FALSE;
        FRealFirst.Bits := DWORD#16#42200000;
        FRealSecond.Bits := DWORD#16#42480000;
        FRealInput[-1] := FRealFirst.Value;
        FRealInput[0] := FRealSecond.Value;
        FRealExpectedFirst := DWORD#16#42200000;
        FRealExpectedSecond := DWORD#16#42480000;
        FLRealFirst.Bits := LWORD#16#4044000000000000;
        FLRealSecond.Bits := LWORD#16#4049000000000000;
        FLRealInput[-1] := FLRealFirst.Value;
        FLRealInput[0] := FLRealSecond.Value;
        FLRealExpectedFirst := LWORD#16#4044000000000000;
        FLRealExpectedSecond := LWORD#16#4049000000000000;
        FRealEnable := TRUE;
        FRealResult := E_Result.NotEvaluated;
        FRealObservation := TRUE;
        FRealEvaluation := FALSE;
        FLRealEnable := TRUE;
        FLRealResult := E_Result.NotEvaluated;
        FLRealObservation := TRUE;
        FLRealEvaluation := FALSE;
    StepCompareNewFinite:
        FTrace := TraceNewSnapshotAfterReset;
        FResetSubjects := FALSE;
        FRealFirst.Bits := DWORD#16#42200000;
        FRealSecond.Bits := DWORD#16#42480000;
        FRealInput[-1] := FRealFirst.Value;
        FRealInput[0] := FRealSecond.Value;
        FRealExpectedFirst := DWORD#16#42200000;
        FRealExpectedSecond := DWORD#16#42480000;
        FLRealFirst.Bits := LWORD#16#4044000000000000;
        FLRealSecond.Bits := LWORD#16#4049000000000000;
        FLRealInput[-1] := FLRealFirst.Value;
        FLRealInput[0] := FLRealSecond.Value;
        FLRealExpectedFirst := LWORD#16#4044000000000000;
        FLRealExpectedSecond := LWORD#16#4049000000000000;
        FRealEnable := TRUE;
        FRealResult := E_Result.Passed;
        FRealObservation := TRUE;
        FRealEvaluation := TRUE;
        FLRealEnable := TRUE;
        FLRealResult := E_Result.Passed;
        FLRealObservation := TRUE;
        FLRealEvaluation := TRUE;
ELSE
    Error(Message := 'Unknown observation checkpoint.');
    RETURN;
END_CASE;
SelectStep := TRUE;
END_METHOD

END_FUNCTION_BLOCK

// ---- Framework/Assertions/POU/Arrays/Real/AssertArrayNoValueChange_Real.TcPOU
{region 'Documentation'}
(*!
<summary>Captures one snapshot until Reset; Disable/Re-Enable never replaces it.</summary>
<description>

Disabling observation preserves the original snapshot. Re-enabling requires a fresh
preceding observation before comparisons resume; it does not replace that snapshot.

StartIndex is an absolute IN index and Length selects 1..255 elements within IN. Memory
must have at least Length elements from its own lower bound. Invalid references or ranges
report Error.

The caller provides dedicated writable Memory that must not overlap IN; overlap is not
checked. Keep bindings, selected range and snapshot contents stable until Reset. Reset
invalidates the snapshot without clearing Memory bytes.

Snapshot capture rejects NaN with Error but accepts either infinity. Later NaN is a
mismatch; equal signed infinities match.

Tolerance is absolute, in the same units as the values, finite and non-negative. Its
default zero requests exact comparison. The equality boundary is inclusive; larger differences
are unequal. Difference checking avoids overflow for large finite operands.

Numeric diagnostics use the formatter's default six significant digits; rounding affects
the message only, not the comparison.

</description>
*)
{endregion}
FUNCTION_BLOCK AssertArrayNoValueChange_Real EXTENDS AssertionBase
VAR_INPUT
    Tolerance : REAL := 0.0; //! Maximum absolute allowed difference; finite and non-negative.
    StartIndex : DINT; //! First selected index in IN; uses the array's declared index range, not a zero-based offset.
    Length : USINT; //! Number of monitored elements, from 1 through 255.
END_VAR
VAR_IN_OUT CONSTANT
    IN : ARRAY[*] OF REAL; //! Read-only actual data; the selected range must remain stable during the call.
END_VAR
VAR_IN_OUT
    Memory : ARRAY[*] OF REAL; //! Dedicated snapshot storage; only this assertion writes its selected elements.
END_VAR
VAR
    FSnapshotValid : BOOL;
    FObservationPrevious : BOOL;
    FEvaluationActive : BOOL;
END_VAR

SUPER^();

